RoboDK station: Vyankatesh_Robotic_Car_Painting_cell.rdk

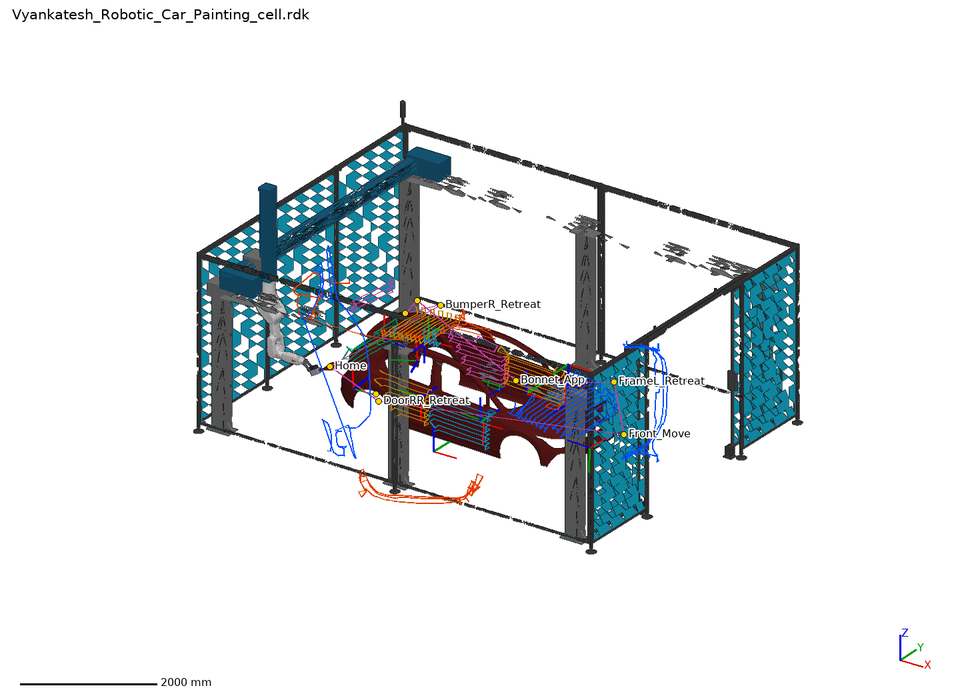
[picture v0: the station drawn from its stored meshes, robots at their saved joint values, targets as dots, program paths as lines]
Station Vyankatesh_Robotic_Car_Painting_cell (saved by RoboDK 6.1.1). Poses are relative to the parent item; angles as X-Y-Z fixed-axis rotations.
Station parameters (name, value as stored): Record_Record, 0, AttachCamera_Record, 0, Surface-Pattern-Generator-Settings, CollisionFreePlanner, ABB IRB 1300-10/1.15, CollisionFreePlanner-Rob ABB IRB 1300-10/1.15
  - frame Frame Car at (0, 0, 0) mm
    - object Trunk_T at (0, 0, 0) mm, size 559.9 x 1436.1 x 749.5 mm, geometry from Trunk_T.stl
    - object Bumper_F_T at (0, 0, 0) mm, size 772.5 x 1766.9 x 440.3 mm, geometry from Bumper_F_T.stl
    - object Bonnet_T at (0, 0, 0) mm, size 1078.9 x 1587.5 x 289.9 mm, geometry from Bonnet_T.stl
    - object Bumper_R_T at (0, 0, 0) mm, size 544.2 x 1726.4 x 536 mm, geometry from Bumper_R_T.stl
    - object Door_FL_T at (0, 0, 0) mm, size 1221.6 x 315.9 x 1113.7 mm, geometry from Door_FL_T.stl
    - object Door_FR_T at (0, 0, 0) mm, size 1221.6 x 316 x 1113.7 mm, geometry from Door_FR_T.stl
    - object Door_RL_T at (0, 0, 0) mm, size 1086.1 x 333.6 x 1090.9 mm, geometry from Door_RL_T.stl
    - object Door_RR_T at (0, 0, 0) mm, size 1086.1 x 333.6 x 1090.9 mm, geometry from Door_RR_T.stl
    - object Frame_T at (0, 0, 0) mm, size 3764.9 x 1786.8 x 1235.6 mm, geometry from Frame_T.stl
    - object Fuel_T at (0, 0, 0) mm, size 294.3 x 103.3 x 136.3 mm, geometry from Fuel_T.stl
    - object Top_T at (0, 0, 0) mm, size 810.7 x 1028.1 x 90.5 mm, geometry from Top_T.stl
    - frame Top2 at (-681.94, -447.22, 1360.45) mm, rotated rx -179.26 ry 1.08 rz -179.99 deg
    - frame Bonnet at (1052.19, 738.82, 942.03) mm, rotated rx 179.6 ry 0.01 rz 1.05 deg
    - frame DoorFL at (817.67, 994, 100.47) mm, rotated rx 105.9 ry -86.47 rz -19.07 deg
      - object DoorFL (SPG) at (0, 0, 0) mm
    - frame DoorRL at (-245.46, 977.17, 107.87) mm, rotated rx 13.73 ry -85.02 rz 76.6 deg
      - object DoorRL (SPG) at (0, 0, 0) mm
    - frame DoorFR at (798.13, -1053.51, 668.15) mm, rotated rx 42.25 ry 86.13 rz 132.32 deg
      - object DoorFR (SPG) at (0, 0, 0) mm
    - frame BumperF at (2280.3, -471.89, 411.2) mm, rotated rx -89.5 ry -0.21 rz 86.56 deg
    - frame DoorRR at (-287.77, -1076.71, 765.51) mm, rotated rx 87.83 ry 88.44 rz 179.37 deg
    - frame Bumper_R at (-1751.94, 908.52, 146.56) mm, rotated rx -73.11 ry -86.07 rz -175.08 deg
    - frame Trunk at (-2141.31, 613.21, 513.17) mm, rotated rx 88.99 ry -89.81 rz 85.05 deg
    - frame FrameL at (-1577.6, 957.23, 510.2) mm, rotated rx 93.66 ry 0 rz 0 deg
      - object FrameL (SPG) at (0, 0, 0) mm
    - frame FrameR at (-1577.79, -967.62, 493.6) mm, rotated rx 8.18 ry -85.7 rz -98.2 deg
      - object FrameR (SPG) at (0, 0, 0) mm
  - frame Cartesian Robot at (0, 0, 0) mm
    - robot My Mechanism: 3 axes
        modified DH rows (alpha deg, a mm, theta deg, d mm): 0, 0, 0, 0 linear; 90, 0, 90, 0 linear; 90, 0, 0, 0 linear
        base shift (0, 0, 0) mm, rotated rx 0 ry -90 rz 180 deg
        joint limits [0, -370, 0] to [5800, 3840, 1100]; home [0, 0, 0]; saved at [0, 0, 0]
      - robot ABB IRB 1300-10/1.15: 6 axes, payload 10 kg, reach 1150 mm, repeatability 0.023 mm, weight 78 kg
          modified DH rows (alpha deg, a mm, theta deg, d mm): 0, 0, 0, 544; -90, 150, -90, 0; 0, 575, 0, 0; -90, 40, 0, 425; 90, 0, 0, 0; -90, 0, 180, 90
          joint limits [-180, -95, -210, -230, -130, -400] to [180, 155, 65, 230, 130, 400]; home [0, 0, 0, 0, 0, 0]; saved at [0, 0, 0, 0, 0, 0]
        - tool Generic Paint Sprayer, TCP at (50, 0, 450) mm, rotated rx 0 ry 30 rz 0 deg, size 277.6 x 203.2 x 501.7 mm
  - frame Frame_Prog at (0, 0, 0) mm
    - target FrameL_Retreat (joint target) at (1421.65, 1379.32, 501.57) mm, rotated rx 178.9 ry 2.61 rz -172.87 deg; joints [31.932, 104.546, -125.413, -151.221, 47.063, 305.481, 2815.734, 3665.468, 738.344] of ABB IRB 1300-10/1.15
    - target Front_Move (Cartesian target) at (2873.26, -440.24, 778.86) mm, rotated rx 124.39 ry -0.68 rz -178.84 deg; joints [-120.26, 86.657, -7.45, -58.906, -114.481, 262.387, 5647.341, 170.911, 1082.66] of ABB IRB 1300-10/1.15
    - target Home (joint target) at (-1449.44, -1750.18, 1201) mm, rotated rx 0 ry -60 rz 180 deg; joints [0, 0, 0, 0, 0, 0, 0, 0, 0] of ABB IRB 1300-10/1.15
    - target BumperR_Retreat (joint target) at (-1695.61, 1414.09, 864.31) mm, rotated rx -107.53 ry 4.62 rz -165.7 deg; joints [-39.158, -91.932, 7.052, 83.863, 76.705, 97.807, 853.022, 3830.081, 364.531] of ABB IRB 1300-10/1.15
    - target Trunk_App (Cartesian target) at (-2045.19, 1025.35, 789.85) mm, rotated rx 93.3 ry 0.38 rz 73.69 deg; joints [-81.249, 102.661, -200.517, 127.066, 82.558, -85.71, 17.635, 2525.27, 659.745] of ABB IRB 1300-10/1.15
    - target Top_Retreat (joint target) at (-1442.79, 464.8, 1389.13) mm, rotated rx -170.97 ry 7.12 rz -173.76 deg; joints [13.22, 135.95, -182.37, -143.59, 7.01, 303.87, 37.44, 2446.95, 0] of ABB IRB 1300-10/1.15
    - target Bonnet_App (joint target) at (1119.24, -686.1, 1265.98) mm, rotated rx 177.3 ry -5.95 rz 179.99 deg; joints [172.493, 123.347, -162.887, -179.232, 74.635, 188.011, 4433.831, 1162.767, 1.741] of ABB IRB 1300-10/1.15
    - target DoorRR_Retreat (joint target) at (-794.82, -1444.65, 696.6) mm, rotated rx 75.81 ry -0.27 rz 178.92 deg; joints [-164.383, 16.979, -25.325, 79.856, 107.569, -167.519, 2238.906, -364.928, 537.904] of ABB IRB 1300-10/1.15
    - target FrameR_App (Cartesian target) at (-1034.25, -1174.19, 640.35) mm, rotated rx 101.61 ry -1.74 rz -171.59 deg; joints [-36.204, 78.94, -160.975, 146.937, -72.367, 90.08, 787.656, -367.42, 482.946] of ABB IRB 1300-10/1.15
  - machining project FrameR: rotZ(0) | rotz(0) | onStart | onPathStart | onApproach | onPoint | onRetract | onFinish | SetRPM(%1) | SetTool(%1) | Extruder(%1) | default | default | OutOnMov(%1) | OutOffMov(%1) | onPathFinish | M_RunCode(%1)
  - machining project FrameL: rotZ(0) | rotz(0) | onStart | onPathStart | onApproach | onPoint | onRetract | onFinish | SetRPM(%1) | SetTool(%1) | Extruder(%1) | default | default | OutOnMov(%1) | OutOffMov(%1) | onPathFinish | M_RunCode(%1)
  - machining project BumperF: rotZ(0) | rotz(0) | onStart | onPathStart | onApproach | onPoint | onRetract | onFinish | SetRPM(%1) | SetTool(%1) | Extruder(%1) | default | default | OutOnMov(%1) | OutOffMov(%1) | onPathFinish | M_RunCode(%1)
  - machining project Bonnet: rotZ(0) | onStart | onPathStart | onApproach | onPoint | onRetract | onFinish | SetRPM(%1) | SetTool(%1) | Extruder(%1) | default | default | OutOnMov(%1) | OutOffMov(%1) | onPathFinish | M_RunCode(%1)
  - machining project Top2: rotZ(0) | rotZ(0) | onStart | onPathStart | onApproach | onPoint | onRetract | onFinish | SetRPM(%1) | SetTool(%1) | Extruder(%1) | default | default | OutOnMov(%1) | OutOffMov(%1) | onPathFinish | M_RunCode(%1)
  - machining project DoorFL: rotZ(0) | rotz(0) | onStart | onPathStart | onApproach | onPoint | onRetract | onFinish | SetRPM(%1) | SetTool(%1) | Extruder(%1) | default | default | OutOnMov(%1) | OutOffMov(%1) | onPathFinish | M_RunCode(%1)
  - machining project DoorRL: rotZ(0) | rotz(0) | onStart | onPathStart | onApproach | onPoint | onRetract | onFinish | SetRPM(%1) | SetTool(%1) | Extruder(%1) | default | default | OutOnMov(%1) | OutOffMov(%1) | onPathFinish | M_RunCode(%1)
  - machining project DoorFR: rotZ(0) | rotZ(0) | onStart | onPathStart | onApproach | onPoint | onRetract | onFinish | SetRPM(%1) | SetTool(%1) | Extruder(%1) | default | default | OutOnMov(%1) | OutOffMov(%1) | onPathFinish | M_RunCode(%1)
  - machining project DoorRR: rotZ(0) | rotz(0) | onStart | onPathStart | onApproach | onPoint | onRetract | onFinish | SetRPM(%1) | SetTool(%1) | Extruder(%1) | default | default | OutOnMov(%1) | OutOffMov(%1) | onPathFinish | M_RunCode(%1)
  - machining project Trunk: rotZ(0) | rotz(0) | onStart | onPathStart | onApproach | onPoint | onRetract | onFinish | SetRPM(%1) | SetTool(%1) | Extruder(%1) | default | default | OutOnMov(%1) | OutOffMov(%1) | onPathFinish | M_RunCode(%1)
  - machining project Bumper_R: rotZ(0) | rotz(0) | onStart | onPathStart | onApproach | onPoint | onRetract | onFinish | SetRPM(%1) | SetTool(%1) | Extruder(%1) | default | default | OutOnMov(%1) | OutOffMov(%1) | onPathFinish | M_RunCode(%1)
  - program Bonnet (314 instructions, listed below)
  - program Top2 (192 instructions, listed below)
  - program DoorRR_C (126 instructions, listed below)
  - program DoorRL_C (142 instructions, listed below)
  - program DoorFL_C (149 instructions, listed below)
  - program DoorFR_C (147 instructions, listed below)
  - program DoorFR (14 instructions, listed below)
  - program BumperR_C (354 instructions, listed below)
  - program Trunk_C (101 instructions, listed below)
  - program Trunk_Top_C (58 instructions, listed below)
  - program Top2_C (192 instructions, listed below)
  - program BumperF (415 instructions, listed below)
  - program BumperF_C (415 instructions, listed below)
  - program FrameL_C (243 instructions, listed below)
  - program FrameR_C (273 instructions, listed below)
  - program Main_Prog (22 instructions, listed below)
  - frame Cell  at (0, 0, 0) mm
    - frame Left at (0, -1180, 0) mm
      - object LeftGlass at (0, 0, 0) mm, size 6 x 1164 x 2469 mm, geometry from LeftGlass.stl
      - object LeftGlassFrame at (0, 0, 0) mm, size 172 x 1253 x 2620 mm, geometry from LeftGlassFrame.stl
    - frame Right at (0, 1180, 0) mm
      - object RightGlass at (0, 0, 0) mm, size 6 x 1166 x 2471 mm, geometry from RightGlass.stl
      - object RightGlassFrame at (0, 0, 0) mm, size 172 x 1253 x 2620 mm, geometry from RightGlassFrame.stl
  - object Floor at (0, 0, 0) mm, size 8000 x 5600 x 0 mm, geometry from Floor.stl
  - object OuterGlass at (0, 0, 0) mm, size 7005.9 x 5255.9 x 2661 mm, geometry from OuterGlass.stl
  - object GlassFrame at (0, 0, 0) mm, size 7159.9 x 5409.9 x 3270 mm, geometry from GlassFrame.stl
  - program DoorRR (126 instructions, listed below)
  - program FrameL (45 instructions, listed below)
  - program FrameR (273 instructions, listed below)
  - program DoorFL (22 instructions, listed below)
  - program DoorRL (15 instructions, listed below)
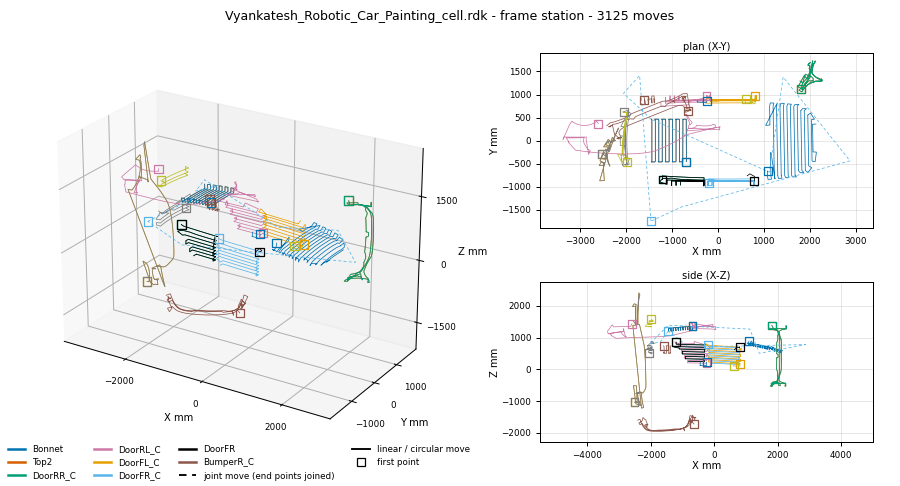
[picture p0: tool path of Vyankatesh_Robotic_Car_Painting_cell.rdk in frame station, 3125 of 3125 moves have a stored position in this frame; points joined in program order, loops and branches not executed]

--- program Bonnet (robot ABB IRB 1300-10/1.15) ---
  Smooth(1)
  Set speed (1000.0 mm/s)
  Set Ref.: Bonnet
  Set Tool: Generic Paint Sprayer
  Show Generic Paint Sprayer
  MoveJ 1 to (13.71, 1405.55, 66.05) mm, rotated rx -3.07 ry 7.94 rz -179.16 deg; joints [173.742, 90.77, -145.127, -180, 57.846, 186.984, 4434.016, 1162.706, 0.414]
  MoveL 2 to (13.71, 1405.55, 66.05) mm, rotated rx -3.07 ry 7.94 rz -179.16 deg; joints [173.742, 90.77, -145.127, -180, 57.846, 186.984, 4434.017, 1162.706, 0.414]
  MoveL 3 to (0, 1400, 164.95) mm, rotated rx -3.07 ry 7.94 rz -179.16 deg; joints [173.742, 90.769, -145.127, -180, 57.846, 186.984, 4420.212, 1167.307, 99.349]
  MoveL 4 to (0, 1400, 164.95) mm, rotated rx -3.07 ry 7.94 rz -179.16 deg; joints [173.742, 90.769, -145.127, -180, 57.846, 186.984, 4420.212, 1167.307, 99.349]
  Set speed (200.0 mm/s)
  MoveL 5 to (0, 1500, 204.66) mm, rotated rx -53.96 ry 9.04 rz 178.26 deg; joints [162.372, 90.769, -145.127, -214.939, 81.944, 234.484, 4381.306, 868.259, 332.309]
  Set speed (1000.0 mm/s)
  MoveL 6 to (0, 1500, 204.66) mm, rotated rx -53.96 ry 9.04 rz 178.26 deg; joints [162.372, 90.769, -145.127, -214.939, 81.944, 234.484, 4381.306, 868.259, 332.309]
  MoveL 7 to (11.7, 1580.54, 146.56) mm, rotated rx -53.96 ry 9.04 rz 178.26 deg; joints [162.372, 90.77, -145.127, -214.939, 81.944, 234.484, 4394.48, 788.358, 273.639]
  Set speed (1000.0 mm/s)
  MoveL 8 to (86.8, 1577.85, 157.52) mm, rotated rx -51.38 ry 9.02 rz 178.52 deg; joints [163.545, 90.769, -145.127, -214.254, 79.866, 232.519, 4475.298, 788.36, 267.392]
  MoveL 9 to (75, 1500, 219.17) mm, rotated rx -51.38 ry 9.02 rz 178.52 deg; joints [163.545, 90.769, -145.127, -214.254, 79.866, 232.519, 4462.081, 865.544, 329.584]
  MoveL 10 to (75, 1500, 219.17) mm, rotated rx -51.38 ry 9.02 rz 178.52 deg; joints [163.545, 90.769, -145.127, -214.254, 79.866, 232.519, 4462.081, 865.544, 329.584]
  Set speed (200.0 mm/s)
  MoveL 11 to (75, 1400, 175.28) mm, rotated rx -2.63 ry 8.05 rz -179.16 deg; joints [163.545, 106.008, -145.127, -175.627, 72.598, 194.93, 4527.686, 1355.214, 329.584]
  MoveL 12 to (75, 1300, 170.07) mm, rotated rx -3.56 ry 8.28 rz -179.19 deg; joints [164.42, 106.008, -145.153, -176.848, 72.598, 194.93, 4532.073, 1432.375, 324.681]
  MoveL 13 to (75, 1200, 162.92) mm, rotated rx -2 ry 7.25 rz -179.12 deg; joints [166.99, 106.008, -145.153, -176.244, 73.416, 191.618, 4532.073, 1502.111, 320.532]
  MoveL 14 to (75, 1100, 159.11) mm, rotated rx -1.73 ry 6.88 rz -179.11 deg; joints [167.767, 106.008, -145.153, -176.244, 73.775, 190.768, 4529.877, 1591.137, 318.443]
  MoveL 15 to (75, 1000, 155.9) mm, rotated rx -1.44 ry 7.2 rz -179.12 deg; joints [167.77, 106.24, -145.152, -176.048, 73.647, 190.576, 4531.483, 1693.74, 318.443]
  Set speed (1000.0 mm/s)
  MoveL 16 to (75, 1000, 155.9) mm, rotated rx -1.44 ry 7.2 rz -179.12 deg; joints [167.77, 106.24, -145.152, -176.048, 73.647, 190.576, 4531.483, 1693.74, 318.443]
  MoveL 17 to (87.48, 1002.7, 56.72) mm, rotated rx -1.44 ry 7.2 rz -179.12 deg; joints [167.77, 106.24, -145.152, -176.048, 73.647, 190.576, 4544.012, 1691.978, 219.247]
  Set speed (1000.0 mm/s)
  MoveL 18 to (163.33, 1574.44, 167.94) mm, rotated rx -44.22 ry 24.07 rz -167.42 deg; joints [161.786, 90.814, -145.127, -206.546, 69.381, 247.678, 4571.543, 889.471, 203.361]
  MoveL 19 to (150, 1500, 233.37) mm, rotated rx -44.22 ry 24.07 rz -167.42 deg; joints [161.786, 90.814, -145.127, -206.546, 69.382, 247.678, 4556.853, 963.186, 269.318]
  MoveL 20 to (150, 1500, 233.37) mm, rotated rx -44.22 ry 24.07 rz -167.42 deg; joints [161.786, 90.814, -145.127, -206.546, 69.382, 247.678, 4556.853, 963.186, 269.318]
  Set speed (200.0 mm/s)
  MoveL 21 to (150, 1400, 185.67) mm, rotated rx 0.71 ry 8.41 rz -158.95 deg; joints [180, 101.307, -145.127, -171.069, 66.652, 194.666, 4644.083, 1152.192, 269.318]
  MoveL 22 to (150, 1300, 180.88) mm, rotated rx -8.15 ry 4.46 rz 140.73 deg; joints [127.726, 83.623, -166.891, -182.813, 33.065, 197.095, 4139.747, 1597.912, 0.019]
  MoveL 23 to (150, 1200, 172.83) mm, rotated rx -2.4 ry 7.56 rz -179.14 deg; joints [25.975, 87.43, -169.901, -43.466, 16.467, 198.768, 2962.972, 1597.586, 18.083]
  MoveL 24 to (150, 1100, 168.79) mm, rotated rx -2.16 ry 7.38 rz -179.13 deg; joints [25.908, 87.621, -170.162, -42.349, 16.618, 197.63, 2959.562, 1698.654, 17.072]
  MoveL 25 to (150, 1000, 165.32) mm, rotated rx -1.64 ry 7.21 rz -179.12 deg; joints [25.707, 87.861, -170.491, -40.208, 16.705, 195.488, 2955.557, 1800.56, 17.072]
  MoveL 26 to (150, 900, 162.41) mm, rotated rx -1.26 ry 7.12 rz -179.12 deg; joints [25.558, 88.036, -170.732, -38.697, 16.743, 193.978, 2952.499, 1901.9, 16.797]
  MoveL 27 to (150, 800, 160.25) mm, rotated rx -1.02 ry 6.68 rz -179.11 deg; joints [25.455, 88.057, -170.76, -37.493, 17.124, 192.798, 2946.147, 2002.771, 16.797]
  MoveL 28 to (150, 700, 159.04) mm, rotated rx 0.41 ry 7.43 rz -179.12 deg; joints [24.734, 88.057, -170.76, -32.755, 16.105, 188.203, 2947.144, 2106.644, 14.156]
  MoveL 29 to (150, 600, 159.34) mm, rotated rx 0.28 ry 6.68 rz -179.12 deg; joints [24.734, 87.748, -170.76, -32.228, 17.13, 187.718, 2940.681, 2204.426, 14.157]
  MoveL 30 to (150, 500, 160.27) mm, rotated rx 0.78 ry 7.01 rz -179.12 deg; joints [24.474, 87.675, -170.719, -30.467, 16.76, 186.011, 2940.681, 2305.628, 14.157]
  MoveL 31 to (150, 400, 161.65) mm, rotated rx 0.99 ry 7.45 rz -179.12 deg; joints [24.363, 87.589, -170.601, -29.905, 16.266, 185.477, 2942.074, 2406.202, 14.157]
  MoveL 32 to (150, 300, 163.74) mm, rotated rx 1.37 ry 7.2 rz -179.12 deg; joints [24.17, 87.589, -170.601, -28.388, 16.481, 184.008, 2936.908, 2507.18, 17.764]
  MoveL 33 to (150, 200, 169.2) mm, rotated rx 2.84 ry 8.35 rz -179.06 deg; joints [23.441, 87.248, -170.135, -23.017, 15.142, 178.814, 2940.939, 2611.654, 17.919]
  MoveL 34 to (150, 100, 172.42) mm, rotated rx 1.6 ry 7.77 rz -179.1 deg; joints [23.441, 86.759, -170.135, -26.264, 16.178, 182.487, 2937.523, 2699.259, 17.919]
  MoveL 35 to (150, 0, 193.42) mm, rotated rx 48.1 ry 9.85 rz -176.1 deg; joints [6.576, 86.759, -170.136, 60.139, 45.852, 96.029, 2889.461, 2951.486, 197.833]
  Set speed (1000.0 mm/s)
  MoveL 36 to (150, 0, 193.42) mm, rotated rx 48.1 ry 9.85 rz -176.1 deg; joints [6.576, 86.759, -170.136, 60.139, 45.852, 96.029, 2889.461, 2951.486, 197.833]
  MoveL 37 to (166.47, -73.48, 127.62) mm, rotated rx 48.1 ry 9.85 rz -176.1 deg; joints [6.576, 86.759, -170.136, 60.139, 45.852, 96.029, 2904.579, 3025.719, 132.557]
  Set speed (1000.0 mm/s)
  MoveL 38 to (89.54, -78.19, 114.09) mm, rotated rx 52.11 ry 9.16 rz -176.52 deg; joints [5.072, 86.759, -170.136, 61.133, 49.725, 94.485, 2815.202, 3031.106, 147.378]
  MoveL 39 to (75, 0, 174.71) mm, rotated rx 52.11 ry 9.16 rz -176.52 deg; joints [5.072, 86.759, -170.136, 61.133, 49.725, 94.486, 2802.092, 2952.242, 207.449]
  MoveL 40 to (75, 0, 174.71) mm, rotated rx 52.11 ry 9.16 rz -176.52 deg; joints [5.072, 86.759, -170.136, 61.133, 49.725, 94.486, 2802.092, 2952.242, 207.449]
  Set speed (200.0 mm/s)
  MoveL 41 to (75, 100, 161.89) mm, rotated rx 1.85 ry 8.11 rz -179.09 deg; joints [23.489, 88.002, -170.136, -27.629, 14.727, 183.787, 2856.802, 2704.635, 19.313]
  MoveL 42 to (75, 200, 158.17) mm, rotated rx 2.73 ry 8.3 rz -179.07 deg; joints [23.489, 88.444, -170.136, -25.354, 14.108, 181.209, 2857.15, 2613.667, 19.312]
  MoveL 43 to (75, 300, 153.75) mm, rotated rx 1.3 ry 7.73 rz -179.11 deg; joints [24.186, 88.444, -170.136, -31.197, 14.806, 186.915, 2857.632, 2509.61, 15.205]
  MoveL 44 to (75, 400, 153.25) mm, rotated rx -65.18 ry 32.47 rz -81.47 deg; joints [-7.384, 82.47, -173.542, 30.828, 55.97, 290.824, 2599.504, 2142.82, 179.665]
  Set speed (1000.0 mm/s)
  MoveL 45 to (75, 400, 153.25) mm, rotated rx -65.18 ry 32.47 rz -81.47 deg; joints [-7.384, 82.47, -173.542, 30.828, 55.97, 290.824, 2599.504, 2142.82, 179.665]
  MoveL 46 to (-18.1, 408.83, 117.84) mm, rotated rx -48.18 ry -57.92 rz -132.58 deg; joints [5.789, 76.051, -169.247, 0, 99.953, 203.081, 2424.003, 2179.227, 396.057]
  Set speed (1000.0 mm/s)
  MoveL 47 to (242.54, -75.07, 148.77) mm, rotated rx 49.67 ry 10.26 rz -175.45 deg; joints [5.789, 76.051, -169.247, 55.04, 52.306, 105.502, 3073.622, 3019.948, 61.16]
  MoveL 48 to (225, 0, 212.46) mm, rotated rx 49.67 ry 10.26 rz -175.45 deg; joints [5.789, 76.051, -169.247, 55.04, 52.306, 105.502, 3057.455, 2944.119, 124.315]
  MoveL 49 to (225, 0, 212.46) mm, rotated rx 49.67 ry 10.26 rz -175.45 deg; joints [5.789, 76.051, -169.247, 55.04, 52.306, 105.502, 3057.455, 2944.119, 124.315]
  Set speed (200.0 mm/s)
  MoveL 50 to (225, 100, 183.39) mm, rotated rx 0.83 ry 8.18 rz -179.11 deg; joints [15.296, 83.487, -177.068, -10.85, 25.36, 174.895, 3057.454, 2574.979, 0]
  MoveL 51 to (225, 200, 180.77) mm, rotated rx 2.66 ry 8.52 rz -179.06 deg; joints [15.296, 83.901, -177.068, -7.153, 24.807, 170.698, 3058.945, 2491.778, 0]
  MoveL 52 to (225, 300, 173.64) mm, rotated rx 1.36 ry 7.35 rz -179.12 deg; joints [15.88, 84.388, -177.768, -10.555, 26.023, 173.843, 3053.064, 2386.704, 0]
  MoveL 53 to (225, 400, 171.5) mm, rotated rx 1.18 ry 7.79 rz -179.11 deg; joints [16.011, 84.85, -177.768, -11.109, 25.117, 174.348, 3055.565, 2287.744, 0]
  MoveL 54 to (225, 500, 169.85) mm, rotated rx 0.84 ry 7.43 rz -179.12 deg; joints [16.182, 84.988, -177.967, -12.016, 25.501, 175.176, 3055.056, 2186.543, 0]
  MoveL 55 to (225, 600, 168.94) mm, rotated rx 0.53 ry 7.14 rz -179.12 deg; joints [16.33, 85.067, -178.08, -12.799, 25.81, 175.895, 3054.866, 2085.487, 0]
  MoveL 56 to (225, 700, 168.3) mm, rotated rx 0.46 ry 7.35 rz -179.12 deg; joints [16.389, 85.287, -178.08, -13.055, 25.373, 176.127, 3057.115, 1986.104, 0]
  MoveL 57 to (225, 800, 169.49) mm, rotated rx -1.24 ry 7.12 rz -179.12 deg; joints [17.175, 85.179, -177.924, -17.239, 25.498, 180.034, 3059.26, 1880.248, 0]
  MoveL 58 to (225, 900, 171.99) mm, rotated rx -1.33 ry 6.99 rz -179.12 deg; joints [17.227, 85.28, -177.924, -17.522, 25.536, 180.297, 3059.26, 1780.347, 3.097]
  MoveL 59 to (225, 1000, 174.93) mm, rotated rx -1.68 ry 7.42 rz -179.13 deg; joints [17.384, 85.177, -177.776, -18.423, 25.066, 181.15, 3065.255, 1679.079, 3.097]
  MoveL 60 to (225, 1100, 178.7) mm, rotated rx -2.17 ry 8.02 rz -179.15 deg; joints [17.597, 85.034, -177.569, -19.725, 24.409, 182.385, 3072.997, 1577.25, 3.097]
  MoveL 61 to (225, 1200, 182.76) mm, rotated rx -2.2 ry 7.73 rz -179.14 deg; joints [17.603, 85.034, -177.569, -19.748, 24.7, 182.411, 3072.215, 1477.151, 7.244]
  MoveL 62 to (225, 1300, 192.42) mm, rotated rx -2.69 ry 8.46 rz -179.18 deg; joints [17.714, 84.444, -176.724, -21.177, 23.751, 183.883, 3079.788, 1374.447, 8.221]
  MoveL 63 to (225, 1400, 196.36) mm, rotated rx -1.65 ry 8.59 rz -179.16 deg; joints [17.714, 84.583, -176.724, -19.035, 23.457, 181.445, 3081.636, 1283.763, 12.105]
  MoveL 64 to (225, 1500, 247.21) mm, rotated rx -41.7 ry 9.43 rz 178.83 deg; joints [27.955, 71.742, -159.319, -88.579, 43.502, 254.167, 3123.032, 976.712, 51.789]
  Set speed (1000.0 mm/s)
  MoveL 65 to (225, 1500, 247.21) mm, rotated rx -41.7 ry 9.43 rz 178.83 deg; joints [27.955, 71.742, -159.319, -88.579, 43.502, 254.167, 3123.032, 976.712, 51.789]
  MoveL 66 to (238.58, 1566.25, 173.55) mm, rotated rx -41.7 ry 9.43 rz 178.83 deg; joints [29.173, 74.127, -159.319, -92.303, 43.597, 257.628, 3123.032, 935.899, 0]
  Set speed (1000.0 mm/s)
  MoveL 67 to (315.52, 1560.78, 183.61) mm, rotated rx -37.7 ry 10.16 rz 178.53 deg; joints [27.986, 75.504, -159.319, -92.621, 39.841, 257.853, 3190.269, 962.686, 0]
  MoveL 68 to (300, 1500, 261.49) mm, rotated rx -37.7 ry 10.16 rz 178.53 deg; joints [27.986, 75.504, -159.319, -92.621, 39.841, 257.853, 3173.641, 1022.617, 78.302]
  MoveL 69 to (300, 1500, 261.49) mm, rotated rx -37.7 ry 10.16 rz 178.53 deg; joints [27.986, 75.504, -159.319, -92.621, 39.841, 257.853, 3173.641, 1022.617, 78.302]
  Set speed (200.0 mm/s)
  MoveL 70 to (300, 1400, 208.07) mm, rotated rx -1.39 ry 8.99 rz -179.17 deg; joints [17.09, 87.326, -175.277, -21.576, 19.105, 184.796, 3126.615, 1290.083, 47.242]
  MoveL 71 to (300, 1300, 204.58) mm, rotated rx -2.31 ry 9.55 rz -179.22 deg; joints [16.15, 87.326, -175.277, -23.211, 18.622, 187.649, 3126.615, 1371.082, 43.238]
  MoveL 72 to (300, 1200, 193.84) mm, rotated rx -2.35 ry 8.91 rz -179.19 deg; joints [16.15, 87.762, -175.895, -22.88, 19.432, 187.336, 3120.036, 1470.451, 39.287]
  MoveL 73 to (300, 1100, 189.49) mm, rotated rx -2.12 ry 8.59 rz -179.17 deg; joints [16.081, 88.023, -176.265, -21.971, 19.824, 186.418, 3115.771, 1571.51, 39.081]
  MoveL 74 to (300, 1000, 185.81) mm, rotated rx -1.83 ry 8.63 rz -179.17 deg; joints [15.939, 88.053, -176.308, -21.088, 19.772, 185.583, 3113.884, 1672.287, 36.248]
  MoveL 75 to (300, 900, 182.49) mm, rotated rx -1.49 ry 8.68 rz -179.16 deg; joints [15.765, 88.088, -176.358, -19.999, 19.711, 184.554, 3111.995, 1773.235, 33.807]
  MoveL 76 to (300, 800, 179.69) mm, rotated rx -1.28 ry 8.26 rz -179.15 deg; joints [15.674, 88.189, -176.502, -19.237, 20.15, 183.816, 3106.38, 1873.929, 33.807]
  MoveL 77 to (300, 700, 178.51) mm, rotated rx 0.42 ry 8.27 rz -179.11 deg; joints [14.803, 88.236, -176.569, -13.977, 20.124, 178.867, 3101.896, 1978.338, 33.807]
  MoveL 78 to (300, 600, 179.27) mm, rotated rx 0.66 ry 8.76 rz -179.1 deg; joints [14.68, 88.216, -176.54, -13.21, 19.632, 178.149, 3104.063, 2078.956, 33.807]
  MoveL 79 to (300, 500, 180.56) mm, rotated rx 1.01 ry 8.7 rz -179.09 deg; joints [14.502, 88.216, -176.54, -12.117, 19.701, 177.121, 3101.147, 2179.85, 36.013]
  MoveL 80 to (300, 400, 182.21) mm, rotated rx 1.26 ry 8.59 rz -179.09 deg; joints [14.374, 88.216, -176.54, -11.346, 19.823, 176.394, 3097.913, 2280.477, 38.718]
  MoveL 81 to (300, 300, 184.43) mm, rotated rx 1.56 ry 9.04 rz -179.07 deg; joints [14.207, 88.036, -176.285, -10.336, 19.316, 175.463, 3099.179, 2381.233, 38.718]
  MoveL 82 to (300, 200, 192.84) mm, rotated rx 2.59 ry 9.4 rz -179.02 deg; joints [13.689, 87.953, -176.21, -6.909, 19.057, 172.229, 3099.179, 2484.02, 46.473]
  MoveL 83 to (300, 100, 194.82) mm, rotated rx 0.83 ry 9.24 rz -179.09 deg; joints [13.689, 87.711, -176.211, -11.528, 19.32, 177.395, 3097.796, 2568.243, 46.707]
  MoveL 84 to (300, 0, 232.6) mm, rotated rx 41.6 ry 10.8 rz -175.86 deg; joints [-6.021, 87.711, -176.211, 68.056, 42.901, 105.13, 3088.96, 2757.637, 205.756]
  Set speed (1000.0 mm/s)
  MoveL 85 to (300, 0, 232.6) mm, rotated rx 41.6 ry 10.8 rz -175.86 deg; joints [-6.021, 87.711, -176.211, 68.056, 42.901, 105.13, 3088.96, 2757.637, 205.756]
  MoveL 86 to (318.77, -65.21, 159.15) mm, rotated rx 41.6 ry 10.8 rz -175.86 deg; joints [-6.021, 87.711, -176.211, 68.056, 42.901, 105.13, 3106.537, 2823.697, 132.769]
  Set speed (1000.0 mm/s)
  MoveL 87 to (394.09, -63.48, 176.58) mm, rotated rx 40.3 ry 10.95 rz -175.88 deg; joints [-5.321, 87.766, -176.211, 67.069, 41.703, 105.865, 3182.413, 2823.062, 143.079]
  MoveL 88 to (375, 0, 251.46) mm, rotated rx 40.3 ry 10.95 rz -175.88 deg; joints [-5.321, 87.766, -176.211, 67.069, 41.703, 105.865, 3164.491, 2758.721, 217.504]
  MoveL 89 to (375, 0, 251.46) mm, rotated rx 40.3 ry 10.95 rz -175.88 deg; joints [-5.321, 87.766, -176.211, 67.069, 41.703, 105.865, 3164.491, 2758.721, 217.504]
  Set speed (200.0 mm/s)
  MoveL 90 to (375, 100, 207.39) mm, rotated rx 0.55 ry 10.1 rz -179.09 deg; joints [13.83, 87.766, -176.211, -12.371, 18.395, 178.193, 3180.679, 2568.934, 57.639]
  MoveL 91 to (375, 200, 205.89) mm, rotated rx 2.6 ry 10.23 rz -178.98 deg; joints [13.83, 88.078, -176.211, -6.727, 18.114, 171.926, 3181.211, 2487.437, 58.72]
  MoveL 92 to (375, 300, 196.95) mm, rotated rx 1.57 ry 9.8 rz -179.05 deg; joints [14.354, 88.197, -176.38, -10.315, 18.496, 175.304, 3181.025, 2384.58, 50.941]
  MoveL 93 to (375, 400, 194.55) mm, rotated rx 1.23 ry 9.65 rz -179.07 deg; joints [14.527, 88.254, -176.38, -11.497, 18.564, 176.419, 3181.65, 2283.834, 48.647]
  MoveL 94 to (375, 500, 192.59) mm, rotated rx 1 ry 9.63 rz -179.08 deg; joints [14.644, 88.254, -176.38, -12.262, 18.582, 177.14, 3183.59, 2183.241, 45.99]
  MoveL 95 to (375, 600, 191.19) mm, rotated rx 0.68 ry 9.25 rz -179.1 deg; joints [14.825, 88.373, -176.549, -13.366, 19, 178.164, 3182.849, 2082.442, 45.99]
  MoveL 96 to (375, 700, 190.31) mm, rotated rx 0.61 ry 9.24 rz -179.1 deg; joints [14.859, 88.373, -176.549, -13.585, 19.005, 178.369, 3184.727, 1982.29, 44.406]
  MoveL 97 to (375, 800, 191.51) mm, rotated rx -1.47 ry 9.25 rz -179.17 deg; joints [15.931, 88.325, -176.482, -20.389, 19.038, 184.772, 3190.004, 1876.825, 44.405]
  MoveL 98 to (375, 900, 194.48) mm, rotated rx -1.72 ry 9.6 rz -179.19 deg; joints [16.032, 88.185, -176.282, -21.327, 18.652, 185.686, 3195.013, 1775.96, 44.405]
  MoveL 99 to (375, 1000, 197.95) mm, rotated rx -1.86 ry 9.61 rz -179.2 deg; joints [16.097, 88.151, -176.234, -21.797, 18.641, 186.135, 3197.071, 1675.545, 46.812]
  MoveL 100 to (375, 1100, 202) mm, rotated rx -2.39 ry 10.09 rz -179.24 deg; joints [16.322, 87.923, -175.91, -23.8, 18.139, 188.075, 3203.415, 1573.734, 46.812]
  MoveL 101 to (375, 1200, 206.54) mm, rotated rx -2.44 ry 9.79 rz -179.23 deg; joints [16.352, 87.923, -175.91, -23.845, 18.441, 188.115, 3202.619, 1473.638, 51.377]
  MoveL 102 to (375, 1300, 217.6) mm, rotated rx -2.03 ry 10.57 rz -179.24 deg; joints [16.352, 87.453, -175.243, -23.259, 17.441, 187.396, 3210.369, 1377.45, 54.97]
  MoveL 103 to (375, 1400, 221) mm, rotated rx -1.2 ry 10.41 rz -179.19 deg; joints [16.352, 87.508, -175.243, -20.821, 17.466, 184.706, 3210.369, 1284.858, 58.398]
  MoveL 104 to (375, 1500, 276.56) mm, rotated rx -29.1 ry 11.25 rz 178.58 deg; joints [25.924, 79.147, -163.83, -87.251, 31.923, 250.899, 3248.664, 1064.43, 86.696]
  Set speed (1000.0 mm/s)
  MoveL 105 to (375, 1500, 276.56) mm, rotated rx -29.1 ry 11.25 rz 178.58 deg; joints [25.924, 79.147, -163.83, -87.251, 31.923, 250.899, 3248.664, 1064.43, 86.696]
  MoveL 106 to (393.24, 1548.2, 190.86) mm, rotated rx -29.1 ry 11.25 rz 178.58 deg; joints [25.924, 79.147, -163.83, -87.251, 31.923, 250.899, 3267.782, 1017.182, 0.665]
  Set speed (1000.0 mm/s)
  MoveL 107 to (470.75, 1541.56, 204.5) mm, rotated rx -24.91 ry 12.47 rz 178.4 deg; joints [24.056, 79.641, -163.83, -85.84, 27.687, 249.752, 3343.92, 1038.3, 0.665]
  MoveL 108 to (450, 1500, 293.05) mm, rotated rx -24.91 ry 12.47 rz 178.4 deg; joints [24.056, 79.64, -163.83, -85.838, 27.687, 249.75, 3322.418, 1078.84, 89.502]
  MoveL 109 to (450, 1500, 293.05) mm, rotated rx -24.91 ry 12.47 rz 178.4 deg; joints [24.056, 79.64, -163.83, -85.838, 27.687, 249.75, 3322.418, 1078.84, 89.502]
  Set speed (200.0 mm/s)
  MoveL 110 to (450, 1400, 235.27) mm, rotated rx -1.57 ry 11.98 rz -179.25 deg; joints [16.298, 86.244, -172.78, -24.148, 14.832, 188.239, 3291.716, 1284.532, 56.208]
  MoveL 111 to (450, 1300, 231.88) mm, rotated rx -2.49 ry 10.96 rz -179.29 deg; joints [16.298, 86.268, -172.814, -26.537, 15.986, 190.936, 3280.502, 1376.523, 56.208]
  MoveL 112 to (450, 1200, 220.89) mm, rotated rx -2.79 ry 11.21 rz -179.32 deg; joints [16.171, 86.268, -172.814, -27.528, 15.785, 192.139, 3280.58, 1472.42, 45.456]
  MoveL 113 to (450, 1100, 215.84) mm, rotated rx -2.44 ry 10.78 rz -179.28 deg; joints [16.073, 86.612, -173.293, -25.8, 16.274, 190.404, 3275.148, 1574.119, 45.456]
  MoveL 114 to (450, 1000, 211.48) mm, rotated rx -2.12 ry 10.68 rz -179.25 deg; joints [15.943, 86.743, -173.476, -24.509, 16.367, 189.139, 3272.269, 1675.333, 43.277]
  MoveL 115 to (450, 900, 207.67) mm, rotated rx -1.59 ry 10.35 rz -179.21 deg; joints [15.732, 86.986, -173.816, -22.34, 16.711, 187.012, 3267.276, 1777.314, 43.277]
  MoveL 116 to (450, 800, 204.58) mm, rotated rx -1.69 ry 10.65 rz -179.22 deg; joints [15.718, 86.986, -173.816, -22.76, 16.419, 187.472, 3268.202, 1876.273, 40.202]
  MoveL 117 to (450, 700, 203.34) mm, rotated rx 0.81 ry 10.66 rz -179.07 deg; joints [14.541, 87.041, -173.892, -13.488, 16.297, 178.578, 3262.711, 1984.048, 40.202]
  MoveL 118 to (450, 600, 204.37) mm, rotated rx 0.72 ry 10.35 rz -179.08 deg; joints [14.542, 86.792, -173.892, -13.596, 16.843, 178.705, 3260.003, 2082.718, 40.219]
  MoveL 119 to (450, 500, 205.98) mm, rotated rx 1.23 ry 10.65 rz -179.04 deg; joints [14.298, 86.674, -173.753, -11.727, 16.545, 176.92, 3260.003, 2184.256, 40.766]
  MoveL 120 to (450, 400, 208.16) mm, rotated rx 1.57 ry 10.79 rz -179.02 deg; joints [14.14, 86.622, -173.753, -10.42, 16.475, 175.664, 3259.369, 2285.216, 42.917]
  MoveL 121 to (450, 300, 210.92) mm, rotated rx 1.89 ry 11.17 rz -178.99 deg; joints [13.984, 86.41, -173.457, -9.176, 16.032, 174.484, 3260.103, 2386.236, 43.472]
  MoveL 122 to (450, 200, 219.9) mm, rotated rx 1.62 ry 10.98 rz -179.01 deg; joints [13.984, 86.209, -173.457, -9.973, 16.397, 175.357, 3258.124, 2483.383, 51.547]
  MoveL 123 to (450, 100, 221.34) mm, rotated rx 0.64 ry 10.9 rz -179.08 deg; joints [13.984, 86.01, -173.457, -12.903, 16.632, 178.582, 3257.11, 2574.411, 51.744]
  MoveL 124 to (450, 0, 270.67) mm, rotated rx 32.3 ry 11.87 rz -176.12 deg; joints [0.856, 86.01, -173.457, 59.201, 33.971, 110.066, 3240.974, 2778.695, 176.115]
  Set speed (1000.0 mm/s)
  MoveL 125 to (450, 0, 270.67) mm, rotated rx 32.3 ry 11.87 rz -176.12 deg; joints [0.856, 86.01, -173.457, 59.201, 33.971, 110.066, 3240.974, 2778.695, 176.115]
  MoveL 126 to (470.95, -52.14, 187.95) mm, rotated rx 32.3 ry 11.87 rz -176.12 deg; joints [0.856, 86.01, -173.457, 59.201, 33.971, 110.066, 3260.969, 2831.795, 93.771]
  Set speed (1000.0 mm/s)
  MoveL 127 to (548.91, -41.08, 202.38) mm, rotated rx 25.21 ry 13.47 rz -176.13 deg; joints [3.891, 86.011, -173.457, 53.673, 27.287, 115.128, 3357.611, 2805.126, 75.591]
  MoveL 128 to (525, 0, 290.36) mm, rotated rx 25.21 ry 13.47 rz -176.13 deg; joints [3.891, 86.011, -173.457, 53.673, 27.287, 115.128, 3334.457, 2762.999, 163.279]
  MoveL 129 to (525, 0, 290.36) mm, rotated rx 25.21 ry 13.47 rz -176.13 deg; joints [3.891, 86.011, -173.457, 53.673, 27.287, 115.128, 3334.457, 2762.999, 163.279]
  Set speed (200.0 mm/s)
  MoveL 130 to (525, 100, 236.85) mm, rotated rx 0.8 ry 12.52 rz -179.04 deg; joints [13.914, 86.011, -173.457, -12.118, 15.008, 177.825, 3346.903, 2576.374, 63.83]
  MoveL 131 to (525, 200, 235.15) mm, rotated rx 1.75 ry 12.7 rz -178.95 deg; joints [13.914, 86.232, -173.457, -8.918, 14.67, 174.354, 3348.601, 2485.185, 63.447]
  MoveL 132 to (525, 300, 226.28) mm, rotated rx 2.21 ry 11.91 rz -178.94 deg; joints [13.914, 86.848, -174.321, -7.561, 15.74, 172.845, 3344.562, 2388.842, 61.889]
  MoveL 133 to (525, 400, 223.05) mm, rotated rx 1.87 ry 11.52 rz -178.98 deg; joints [14.083, 87.066, -174.626, -8.951, 16.19, 174.159, 3343.766, 2287.769, 60.885]
  MoveL 134 to (525, 500, 220.45) mm, rotated rx 1.32 ry 11.15 rz -179.03 deg; joints [14.354, 87.225, -174.85, -11.057, 16.584, 176.157, 3343.429, 2186.069, 59.85]
  MoveL 135 to (525, 600, 218.67) mm, rotated rx 0.9 ry 11.04 rz -179.06 deg; joints [14.552, 87.229, -174.85, -12.593, 16.671, 177.622, 3344.831, 2084.81, 57.555]
  MoveL 136 to (525, 700, 217.56) mm, rotated rx 0.68 ry 11 rz -179.07 deg; joints [14.658, 87.229, -174.85, -13.411, 16.7, 178.402, 3346.683, 1984.14, 55.774]
  MoveL 137 to (525, 800, 218.74) mm, rotated rx -1.55 ry 11 rz -179.23 deg; joints [15.727, 87.181, -174.782, -21.522, 16.778, 186.136, 3351.822, 1877.282, 55.774]
  MoveL 138 to (525, 900, 222) mm, rotated rx -1.77 ry 11.02 rz -179.24 deg; joints [15.823, 87.122, -174.699, -22.333, 16.753, 186.918, 3354.061, 1776.55, 57.713]
  MoveL 139 to (525, 1000, 226.01) mm, rotated rx -2.21 ry 11.97 rz -179.31 deg; joints [16.001, 86.988, -174.511, -24.429, 15.823, 188.951, 3364.872, 1674.895, 57.712]
  MoveL 140 to (525, 1100, 230.94) mm, rotated rx -2.79 ry 12.13 rz -179.37 deg; joints [16.238, 86.76, -174.191, -26.832, 15.669, 191.292, 3368.51, 1572.716, 59.455]
  MoveL 141 to (525, 1200, 236.47) mm, rotated rx -3.19 ry 12.26 rz -179.41 deg; joints [16.395, 86.595, -173.959, -28.507, 15.564, 192.93, 3371.66, 1471.164, 62.491]
  MoveL 142 to (525, 1300, 247.7) mm, rotated rx -2.64 ry 12.69 rz -179.38 deg; joints [16.395, 86.387, -173.668, -27.141, 14.968, 191.393, 3376.989, 1376.085, 69.84]
  MoveL 143 to (525, 1400, 251.45) mm, rotated rx -1.65 ry 12.56 rz -179.28 deg; joints [16.395, 86.473, -173.668, -23.827, 14.87, 187.799, 3376.99, 1284.918, 73.706]
  MoveL 144 to (525, 1500, 311.34) mm, rotated rx -22.15 ry 13.64 rz 178.22 deg; joints [23.268, 80.36, -165.33, -83.718, 24.867, 247.081, 3409.347, 1091.269, 103.416]
  Set speed (1000.0 mm/s)
  MoveL 145 to (525, 1500, 311.34) mm, rotated rx -22.15 ry 13.64 rz 178.22 deg; joints [23.268, 80.36, -165.33, -83.718, 24.867, 247.081, 3409.347, 1091.269, 103.416]
  MoveL 146 to (548, 1537.02, 221.34) mm, rotated rx -22.15 ry 13.64 rz 178.22 deg; joints [23.268, 80.36, -165.33, -83.719, 24.867, 247.081, 3433.018, 1055.316, 13.155]
  Set speed (1000.0 mm/s)
  MoveL 147 to (628.79, 1537.21, 244.37) mm, rotated rx -22.8 ry 16.82 rz 176.81 deg; joints [23.268, 78.379, -162.701, -93.295, 24.002, 256.17, 3544.956, 1051.311, 13.155]
  MoveL 148 to (600, 1500, 332.61) mm, rotated rx -22.8 ry 16.82 rz 176.81 deg; joints [23.268, 78.379, -162.701, -93.295, 24.002, 256.17, 3515.485, 1087.363, 101.652]
  MoveL 149 to (600, 1500, 332.61) mm, rotated rx -22.8 ry 16.82 rz 176.81 deg; joints [23.268, 78.379, -162.701, -93.295, 24.002, 256.17, 3515.485, 1087.363, 101.652]
  Set speed (200.0 mm/s)
  MoveL 150 to (600, 1400, 274.62) mm, rotated rx -53.63 ry 16.6 rz 168.42 deg; joints [23.268, 68.229, -149.644, -107.057, 52.228, 277.868, 3548.034, 964.026, 101.652]
  MoveL 151 to (600, 1300, 265.21) mm, rotated rx -2.11 ry 13.55 rz -179.36 deg; joints [15.353, 87.464, -175.061, -24.153, 14.305, 189.25, 3458.118, 1369.187, 96.492]
  MoveL 152 to (600, 1200, 253.06) mm, rotated rx -3.19 ry 12.8 rz -179.44 deg; joints [15.353, 87.812, -175.553, -27.137, 15.346, 192.555, 3450.308, 1459.46, 90.351]
  MoveL 153 to (600, 1100, 247.23) mm, rotated rx -3.04 ry 12.84 rz -179.42 deg; joints [15.275, 87.816, -175.559, -26.56, 15.282, 192.01, 3448.571, 1559.918, 85.14]
  MoveL 154 to (600, 1000, 242.06) mm, rotated rx -2.71 ry 13.21 rz -179.41 deg; joints [15.1, 87.816, -175.559, -25.512, 14.856, 191.031, 3449.625, 1660.776, 79.841]
  MoveL 155 to (600, 900, 237.87) mm, rotated rx -1.89 ry 13.57 rz -179.33 deg; joints [14.684, 87.816, -175.559, -22.386, 14.371, 188.079, 3449.844, 1763.078, 75.457]
  MoveL 156 to (600, 800, 234.49) mm, rotated rx -1.57 ry 11.97 rz -179.25 deg; joints [14.557, 87.816, -175.559, -20.432, 15.929, 186.188, 3432.765, 1864.372, 75.856]
  MoveL 157 to (600, 700, 233.33) mm, rotated rx 0.69 ry 11.98 rz -179.06 deg; joints [13.447, 87.864, -175.627, -11.79, 15.85, 177.982, 3427.852, 1970.986, 75.856]
  MoveL 158 to (600, 600, 234.48) mm, rotated rx 0.95 ry 12.01 rz -179.04 deg; joints [13.321, 87.864, -175.627, -10.798, 15.833, 177.039, 3425.9, 2071.723, 77.709]
  MoveL 159 to (600, 500, 236.34) mm, rotated rx 1.33 ry 12.06 rz -179.01 deg; joints [13.134, 87.864, -175.627, -9.323, 15.8, 175.638, 3424.022, 2172.825, 80.254]
  MoveL 160 to (600, 400, 239.22) mm, rotated rx 2.13 ry 12.08 rz -178.94 deg; joints [12.748, 87.864, -175.627, -6.291, 15.852, 172.755, 3421.253, 2275.163, 84.05]
  MoveL 161 to (600, 300, 242.78) mm, rotated rx 2.3 ry 12.82 rz -178.89 deg; joints [12.65, 87.584, -175.231, -5.297, 15.024, 171.826, 3425.246, 2375.681, 84.05]
  MoveL 162 to (600, 200, 252.4) mm, rotated rx 2.38 ry 13.75 rz -178.84 deg; joints [12.588, 86.947, -174.335, -4.514, 13.848, 171.106, 3430.34, 2475.951, 86.178]
  MoveL 163 to (600, 100, 254.03) mm, rotated rx 0.9 ry 13.96 rz -179.01 deg; joints [12.588, 86.797, -174.156, -10.053, 13.482, 177.062, 3430.34, 2562.923, 86.178]
  MoveL 164 to (600, 0, 311.59) mm, rotated rx 22.65 ry 15.9 rz -175.46 deg; joints [3.252, 86.797, -174.156, 57.28, 23.905, 113.435, 3432.163, 2736.265, 179.12]
  Set speed (1000.0 mm/s)
  MoveL 165 to (600, 0, 311.59) mm, rotated rx 22.65 ry 15.9 rz -175.46 deg; joints [3.252, 86.797, -174.156, 57.28, 23.905, 113.435, 3432.163, 2736.265, 179.12]
  MoveL 166 to (628.25, -36.39, 222.83) mm, rotated rx 22.65 ry 15.9 rz -175.46 deg; joints [3.252, 86.797, -174.156, 57.281, 23.905, 113.435, 3459.739, 2773.788, 90.624]
  Set speed (1000.0 mm/s)
  MoveL 167 to (712.58, -33.86, 251.33) mm, rotated rx 22.3 ry 21.19 rz -173.41 deg; joints [3.686, 84.732, -171.286, 72.055, 20.986, 99.405, 3593.386, 2773.788, 90.624]
  MoveL 168 to (675, 0, 337.6) mm, rotated rx 22.3 ry 21.19 rz -173.41 deg; joints [3.686, 84.732, -171.286, 72.055, 20.986, 99.405, 3556.436, 2738.642, 176.644]
  MoveL 169 to (675, 0, 337.6) mm, rotated rx 22.3 ry 21.19 rz -173.41 deg; joints [3.686, 84.732, -171.286, 72.055, 20.986, 99.405, 3556.436, 2738.642, 176.644]
  Set speed (200.0 mm/s)
  MoveL 170 to (675, 100, 289.19) mm, rotated rx 39.45 ry 19.85 rz -168.87 deg; joints [1.08, 84.732, -171.286, 79.758, 36.632, 90.838, 3557.37, 2738.642, 200.588]
  MoveL 171 to (675, 200, 272.28) mm, rotated rx 1.72 ry 16.92 rz -178.83 deg; joints [14.445, 85.619, -172.512, -7.866, 10.146, 172.848, 3537.533, 2494.458, 87.48]
  MoveL 172 to (675, 300, 263.14) mm, rotated rx 25.19 ry 17.48 rz -174.27 deg; joints [6.222, 84.677, -172.512, 59.363, 25.343, 108.29, 3537.533, 2494.458, 113.755]
  MoveL 173 to (675, 400, 257.86) mm, rotated rx 2.09 ry 16.04 rz -178.79 deg; joints [14.646, 84.678, -172.512, -6.397, 12, 171.061, 3541.097, 2298.24, 63.888]
  MoveL 174 to (675, 500, 254.88) mm, rotated rx 1.86 ry 14.69 rz -178.87 deg; joints [14.751, 84.844, -172.743, -8.235, 13.377, 172.829, 3530.949, 2197.341, 63.889]
  MoveL 175 to (675, 600, 253.18) mm, rotated rx 0.89 ry 14.98 rz -179 deg; joints [15.147, 84.844, -172.743, -12.404, 13.014, 176.866, 3536.758, 2093.484, 60.761]
  MoveL 176 to (675, 700, 252.08) mm, rotated rx 0.84 ry 14.94 rz -179.01 deg; joints [15.17, 84.866, -172.743, -12.676, 13.027, 177.129, 3538.133, 1993.359, 59.215]
  MoveL 177 to (675, 800, 253.29) mm, rotated rx -1.74 ry 14.93 rz -179.36 deg; joints [16.235, 84.815, -172.671, -24.182, 13.134, 188.258, 3543.375, 1883.209, 59.215]
  MoveL 178 to (675, 900, 256.88) mm, rotated rx -1.85 ry 16.51 rz -179.42 deg; joints [16.247, 84.758, -172.592, -25.821, 11.568, 189.885, 3559.914, 1782.421, 59.215]
  MoveL 179 to (675, 1000, 261.11) mm, rotated rx -2.87 ry 16.28 rz -179.58 deg; joints [16.672, 84.708, -172.523, -30.576, 11.97, 194.481, 3561.034, 1678.383, 62.826]
  MoveL 180 to (675, 1100, 266.53) mm, rotated rx -2.99 ry 16.02 rz -179.59 deg; joints [16.728, 84.708, -172.523, -30.832, 12.255, 194.719, 3560.583, 1577.965, 67.954]
  MoveL 181 to (675, 1200, 275.83) mm, rotated rx -22.66 ry 17.79 rz 176.44 deg; joints [23.548, 80.666, -167.003, -91.299, 23.442, 253.196, 3606.044, 1389.3, 67.954]
  MoveL 182 to (675, 1300, 286.17) mm, rotated rx -2.35 ry 16.54 rz -179.51 deg; joints [17.144, 82.999, -170.168, -30.734, 11.062, 194.062, 3567.724, 1389.3, 67.954]
  MoveL 183 to (675, 1400, 310.92) mm, rotated rx -32.35 ry 21.64 rz 171.85 deg; joints [23.561, 74.061, -158.292, -109.263, 31.238, 272.436, 3655.744, 1115.534, 67.954]
  Set speed (1000.0 mm/s)
  MoveL 184 to (675, 1400, 310.92) mm, rotated rx -32.35 ry 21.64 rz 171.85 deg; joints [23.561, 74.061, -158.292, -109.263, 31.238, 272.436, 3655.744, 1115.534, 67.954]
  MoveL 185 to (713.42, 1448.55, 232.39) mm, rotated rx -32.35 ry 21.64 rz 171.85 deg; joints [24.253, 75.281, -158.292, -111.772, 31.737, 274.571, 3687.267, 1081.103, 1.051]
  Set speed (1000.0 mm/s)
  MoveL 186 to (791.32, 1441.6, 268.91) mm, rotated rx -27.86 ry 23.6 rz 172.33 deg; joints [22.471, 75.281, -158.292, -114.054, 27.303, 277.175, 3772.507, 1105.567, 18.49]
  MoveL 187 to (750, 1400, 349.92) mm, rotated rx -27.86 ry 23.6 rz 172.33 deg; joints [20.4, 70.83, -158.292, -103.642, 25.698, 267.854, 3764.211, 1105.567, 57.429]
  MoveL 188 to (750, 1400, 349.92) mm, rotated rx -27.86 ry 23.6 rz 172.33 deg; joints [20.4, 70.83, -158.292, -103.642, 25.698, 267.854, 3764.211, 1105.567, 57.429]
  Set speed (200.0 mm/s)
  MoveL 189 to (750, 1300, 312.16) mm, rotated rx -2.71 ry 20.61 rz -179.76 deg; joints [16.885, 79.551, -169.871, -28.548, 9.89, 191.975, 3707.54, 1376.214, 57.429]
  MoveL 190 to (750, 1200, 303.7) mm, rotated rx -10.82 ry 20.92 rz 178.25 deg; joints [16.885, 79.551, -169.871, -62.155, 13.172, 227.09, 3709.968, 1405.79, 56.641]
  MoveL 191 to (750, 1100, 291.11) mm, rotated rx -3.1 ry 20.44 rz -179.84 deg; joints [14.642, 81.376, -172.383, -26.442, 10.742, 192.162, 3697.195, 1547.027, 56.641]
  MoveL 192 to (750, 1000, 285.42) mm, rotated rx -2.86 ry 20.75 rz -179.8 deg; joints [14.551, 81.376, -172.383, -25.502, 10.398, 191.262, 3697.99, 1648.165, 51.356]
  MoveL 193 to (750, 900, 280.81) mm, rotated rx -1.98 ry 21.15 rz -179.6 deg; joints [14.24, 81.376, -172.383, -21.065, 9.883, 186.968, 3698.994, 1752.406, 46.962]
  MoveL 194 to (750, 800, 277.21) mm, rotated rx -1.38 ry 18.58 rz -179.4 deg; joints [14.09, 81.468, -172.51, -17.056, 12.444, 183.019, 3672.53, 1855.728, 46.962]
  MoveL 195 to (750, 700, 275.91) mm, rotated rx 0.44 ry 18.58 rz -179.03 deg; joints [13.465, 81.526, -172.591, -8.804, 12.499, 175.017, 3668.988, 1964.658, 46.962]
  MoveL 196 to (750, 600, 276.71) mm, rotated rx 0.93 ry 18.76 rz -178.93 deg; joints [13.297, 81.456, -172.585, -6.493, 12.427, 172.777, 3668.988, 2066.864, 47.715]
  MoveL 197 to (750, 500, 278.49) mm, rotated rx 1.89 ry 18.63 rz -178.74 deg; joints [12.973, 81.455, -172.585, -2.328, 12.698, 168.738, 3665.03, 2171.614, 50.583]
  MoveL 198 to (750, 400, 281.44) mm, rotated rx 2.15 ry 20.48 rz -178.62 deg; joints [12.878, 81.244, -172.292, 0.767, 10.854, 165.734, 3680.133, 2272.784, 50.583]
  MoveL 199 to (750, 300, 291.13) mm, rotated rx 9.87 ry 21 rz -176.72 deg; joints [10.471, 81.243, -172.292, 33.174, 13.802, 134.358, 3678.246, 2412.156, 67.586]
  MoveL 200 to (750, 200, 296.86) mm, rotated rx 1.74 ry 20.62 rz -178.71 deg; joints [10.471, 80.549, -172.292, 1.116, 11.328, 167.876, 3678.241, 2440.362, 60.907]
  MoveL 201 to (750, 100, 327.89) mm, rotated rx 31.34 ry 23.33 rz -169.47 deg; joints [2.918, 79.231, -170.474, 74.299, 29.403, 98.188, 3704.792, 2697.231, 145.455]
  Set speed (1000.0 mm/s)
  MoveL 202 to (750, 100, 327.89) mm, rotated rx 31.34 ry 23.33 rz -169.47 deg; joints [2.918, 79.231, -170.474, 74.299, 29.403, 98.188, 3704.792, 2697.231, 145.455]
  MoveL 203 to (792.76, 55.05, 249.46) mm, rotated rx 31.34 ry 23.33 rz -169.47 deg; joints [2.918, 79.231, -170.474, 74.299, 29.403, 98.187, 3746.723, 2743.509, 67.352]
  Set speed (1000.0 mm/s)
  MoveL 204 to (875.06, 62.02, 294.05) mm, rotated rx 28.27 ry 27.97 rz -168.28 deg; joints [5.851, 76.163, -166.316, 82.951, 25.17, 87.992, 3875.398, 2741.042, 67.352]
  MoveL 205 to (825, 100, 371.84) mm, rotated rx 28.27 ry 27.97 rz -168.28 deg; joints [5.851, 76.163, -166.316, 82.951, 25.17, 87.992, 3826.037, 2701.608, 144.865]
  MoveL 206 to (825, 100, 371.84) mm, rotated rx 28.27 ry 27.97 rz -168.28 deg; joints [5.851, 76.163, -166.316, 82.951, 25.17, 87.992, 3826.037, 2701.608, 144.865]
  Set speed (200.0 mm/s)
  MoveL 207 to (825, 200, 327.16) mm, rotated rx 2.48 ry 23.88 rz -178.4 deg; joints [10.291, 78.434, -169.385, 11.215, 7.587, 157.912, 3781.731, 2446.04, 68.575]
  MoveL 208 to (825, 300, 322.5) mm, rotated rx 4.92 ry 24.58 rz -177.63 deg; joints [10.292, 78.434, -169.385, 27.797, 8.058, 140.984, 3790.367, 2367.041, 64.537]
  MoveL 209 to (825, 400, 311.37) mm, rotated rx 2.47 ry 24.85 rz -178.36 deg; joints [10.887, 79.034, -169.385, 15.039, 6.103, 153.51, 3790.387, 2253.95, 56.759]
  MoveL 210 to (825, 500, 308.31) mm, rotated rx 1.97 ry 24.92 rz -178.51 deg; joints [11.012, 79.326, -169.385, 11.823, 5.577, 156.676, 3790.424, 2151.643, 55.479]
  MoveL 211 to (825, 600, 306.59) mm, rotated rx 0.92 ry 22.95 rz -178.87 deg; joints [11.32, 79.567, -169.714, -1.525, 7.305, 169.853, 3774.482, 2046.202, 55.479]
  MoveL 212 to (825, 700, 305.89) mm, rotated rx 0.51 ry 22.75 rz -178.98 deg; joints [11.44, 79.665, -169.807, -4.742, 7.446, 173.018, 3774.482, 1944.063, 55.029]
  MoveL 213 to (825, 800, 307.3) mm, rotated rx -1.49 ry 22.73 rz -179.52 deg; joints [12.012, 79.594, -169.711, -19.257, 7.435, 187.307, 3777.558, 1833.335, 55.029]
  MoveL 214 to (825, 900, 311.14) mm, rotated rx -2.06 ry 25.2 rz -179.76 deg; joints [12.106, 79.304, -169.315, -28.871, 5.008, 196.89, 3802.825, 1729.83, 55.029]
  MoveL 215 to (825, 1000, 315.93) mm, rotated rx -2.98 ry 24.9 rz 179.96 deg; joints [12.372, 79.304, -169.315, -36.424, 5.577, 204.324, 3802.502, 1624.918, 59.358]
  MoveL 216 to (825, 1100, 322.07) mm, rotated rx -3.49 ry 24.81 rz 179.81 deg; joints [12.517, 79.285, -169.289, -40.401, 5.845, 208.237, 3803.934, 1522.16, 64.788]
  MoveL 217 to (825, 1200, 336.02) mm, rotated rx -6.42 ry 24.3 rz 178.96 deg; joints [13.358, 79.144, -169.154, -56.973, 7.787, 224.446, 3803.934, 1406.373, 78.47]
  MoveL 218 to (825, 1300, 343.92) mm, rotated rx -3.79 ry 26.61 rz 179.6 deg; joints [13.358, 78.57, -168.375, -56.934, 4.369, 223.926, 3826.812, 1329.569, 78.47]
  MoveL 219 to (825, 1400, 396.1) mm, rotated rx -32.35 ry 30.71 rz 166.68 deg; joints [15.329, 68.432, -155.051, -118.568, 28.899, 286.323, 3903.548, 1030.981, 96.942]
  Set speed (1000.0 mm/s)
  MoveL 220 to (825, 1400, 396.1) mm, rotated rx -32.35 ry 30.71 rz 166.68 deg; joints [15.329, 68.432, -155.051, -118.568, 28.899, 286.323, 3903.548, 1030.981, 96.942]
  MoveL 221 to (879.31, 1442.13, 323.47) mm, rotated rx -32.35 ry 30.71 rz 166.68 deg; joints [17.436, 73.73, -155.051, -128.002, 31.999, 294.825, 3911.486, 1030.981, 74.748]
  Set speed (1000.0 mm/s)
  MoveL 222 to (965.01, 1345.04, 338.67) mm, rotated rx -41.13 ry 35.66 rz 158.45 deg; joints [14.272, 67.774, -147.513, -134.75, 40.963, 303.605, 4063.849, 1052.925, 74.748]
  MoveL 223 to (900, 1300, 399.87) mm, rotated rx -41.13 ry 35.66 rz 158.45 deg; joints [12.661, 61.615, -147.513, -127.551, 36.751, 296.423, 4063.819, 1060.857, 78.96]
  MoveL 224 to (900, 1300, 399.87) mm, rotated rx -41.13 ry 35.66 rz 158.45 deg; joints [12.661, 61.615, -147.513, -127.551, 36.751, 296.423, 4063.819, 1060.857, 78.96]
  Set speed (200.0 mm/s)
  MoveL 225 to (900, 1200, 376.45) mm, rotated rx -5.76 ry 30.98 rz 178.53 deg; joints [12.661, 74.813, -164.49, -119.412, 4.813, 287.169, 3947.418, 1406.267, 78.96]
  MoveL 226 to (900, 1100, 361.42) mm, rotated rx -3.92 ry 32.3 rz 179.2 deg; joints [12.288, 74.813, -164.49, -143.989, 3.996, 311.895, 3956.588, 1517.577, 65.08]
  MoveL 227 to (900, 1000, 354.79) mm, rotated rx -14.05 ry 26.9 rz 157.11 deg; joints [-32.272, 78.235, -200.496, -17.821, 39, 209.606, 4213.787, 1161.862, 187.031]
  MoveL 228 to (900, 900, 349.34) mm, rotated rx -13.2 ry 27.48 rz 157.37 deg; joints [-32.375, 78.085, -200.64, -16.957, 38.461, 208.928, 4216.39, 1270.934, 180.861]
  MoveL 229 to (900, 800, 345.1) mm, rotated rx -13.01 ry 27.67 rz 157.42 deg; joints [-32.401, 78.017, -200.705, -16.771, 38.353, 208.78, 4216.459, 1373.421, 177.028]
  MoveL 230 to (900, 700, 343.45) mm, rotated rx -10.57 ry 28.58 rz 158.28 deg; joints [-32.624, 77.999, -200.723, -14.06, 36.727, 206.63, 4216.181, 1494.123, 172.897]
  MoveL 231 to (900, 600, 344.2) mm, rotated rx -9.9 ry 28.75 rz 158.52 deg; joints [-32.683, 78.04, -200.684, -13.268, 36.278, 205.994, 4213.532, 1599.163, 173.622]
  MoveL 232 to (900, 500, 346.25) mm, rotated rx 2.21 ry 29.82 rz -178.26 deg; joints [11.263, 75.247, -165.781, 62.747, 2.525, 105.588, 3924.669, 2154.676, 56.079]
  MoveL 233 to (900, 400, 349.42) mm, rotated rx 2.52 ry 29.79 rz -178.14 deg; joints [11.22, 75.019, -165.781, 59.596, 2.898, 108.755, 3924.668, 2256.231, 57.992]
  MoveL 234 to (900, 300, 360.64) mm, rotated rx 4 ry 28.77 rz -177.63 deg; joints [11.046, 73.835, -165.781, 42.791, 5.29, 125.576, 3924.668, 2364.389, 59.462]
  MoveL 235 to (900, 200, 375.7) mm, rotated rx 36.02 ry 33.05 rz -161.56 deg; joints [9.544, 70.977, -161.993, 91.85, 31.049, 77.003, 3995.671, 2681.475, 130.978]
  Set speed (1000.0 mm/s)
  MoveL 236 to (900, 200, 375.7) mm, rotated rx 36.02 ry 33.05 rz -161.56 deg; joints [9.544, 70.977, -161.993, 91.85, 31.049, 77.003, 3995.671, 2681.475, 130.978]
  MoveL 237 to (960.45, 158.17, 307.9) mm, rotated rx 36.02 ry 33.05 rz -161.56 deg; joints [9.544, 70.977, -161.993, 91.85, 31.049, 77.002, 4055.342, 2724.88, 63.491]
  Set speed (1000.0 mm/s)
  MoveL 238 to (1041.93, 291.42, 339.37) mm, rotated rx 8.94 ry 41.66 rz -173.99 deg; joints [10.264, 74.058, -161.993, 143.618, 15.526, 25.688, 4156.509, 2401.707, 63.491]
  MoveL 239 to (975, 300, 413.17) mm, rotated rx 8.94 ry 41.66 rz -173.99 deg; joints [10.264, 74.058, -161.993, 143.618, 15.526, 25.688, 4089.748, 2391.385, 137.221]
  MoveL 240 to (975, 300, 413.17) mm, rotated rx 8.94 ry 41.66 rz -173.99 deg; joints [10.264, 74.058, -161.993, 143.618, 15.526, 25.688, 4089.748, 2391.385, 137.221]
  Set speed (200.0 mm/s)
  MoveL 241 to (975, 400, 400.41) mm, rotated rx 4.06 ry 41.94 rz -176.78 deg; joints [10.774, 74.44, -161.993, 157.274, 14.713, 11.644, 4089.749, 2264.031, 124.28]
  MoveL 242 to (975, 500, 396.79) mm, rotated rx 2.59 ry 38.7 rz -177.76 deg; joints [10.961, 75.781, -163.762, 157.971, 10.9, 10.759, 4061.919, 2157.086, 124.28]
  MoveL 243 to (975, 600, 394.59) mm, rotated rx 1.93 ry 38.54 rz -178.11 deg; joints [11.066, 75.847, -163.778, 160.531, 10.693, 8.123, 4061.919, 2053.636, 121.425]
  MoveL 244 to (975, 700, 393.54) mm, rotated rx 1.21 ry 38.77 rz -178.48 deg; joints [11.162, 75.996, -163.778, 163.856, 10.995, 4.739, 4064.622, 1949.682, 121.424]
  MoveL 245 to (975, 800, 395.49) mm, rotated rx -2.48 ry 38.78 rz 179.57 deg; joints [11.767, 75.861, -163.599, 178.471, 11.194, -10.287, 4068.109, 1829.555, 121.424]
  MoveL 246 to (975, 900, 400.77) mm, rotated rx -3.18 ry 38.51 rz 179.21 deg; joints [11.898, 75.861, -163.599, 181.467, 11.062, -13.371, 4067.93, 1725.804, 125.589]
  MoveL 247 to (975, 1000, 407.69) mm, rotated rx -4.42 ry 41.61 rz 178.35 deg; joints [11.898, 74.393, -161.663, 181.713, 14.768, -13.651, 4098.624, 1618.252, 125.589]
  MoveL 248 to (975, 1100, 416.35) mm, rotated rx -5.44 ry 41.77 rz 177.76 deg; joints [12.017, 74.125, -161.311, 184.206, 15.239, -16.235, 4102.627, 1512.579, 131.886]
  MoveL 249 to (975, 1200, 433.48) mm, rotated rx -10.6 ry 42.1 rz 174.72 deg; joints [12.562, 73.019, -159.867, 195.218, 17.612, -27.654, 4111.909, 1383.404, 142.831]
  Set speed (1000.0 mm/s)
  MoveL 250 to (975, 1200, 433.48) mm, rotated rx -10.6 ry 42.1 rz 174.72 deg; joints [12.562, 73.019, -159.867, 195.218, 17.612, -27.654, 4111.909, 1383.404, 142.831]
  MoveL 251 to (1042.32, 1212.25, 360.55) mm, rotated rx -10.6 ry 42.1 rz 174.72 deg; joints [12.833, 76.294, -159.867, 192.739, 20.795, -25.317, 4147.888, 1383.404, 101.263]
  Set speed (1000.0 mm/s)
  MoveL 252 to (1072.23, 1006.4, 362.98) mm, rotated rx -5.62 ry 46.22 rz 177.3 deg; joints [11.712, 75, -158.186, 180.212, 23.524, -12.101, 4205.736, 1613.499, 101.263]
  MoveL 253 to (1000, 1000, 431.84) mm, rotated rx -5.62 ry 46.22 rz 177.3 deg; joints [11.709, 72.808, -158.186, 180.236, 21.333, -12.122, 4155.35, 1613.499, 148.926]
  MoveL 254 to (1000, 1000, 431.84) mm, rotated rx -5.62 ry 46.22 rz 177.3 deg; joints [11.709, 72.808, -158.186, 180.236, 21.333, -12.122, 4155.35, 1613.499, 148.926]
  Set speed (200.0 mm/s)
  MoveL 255 to (1000, 900, 423.58) mm, rotated rx -4.13 ry 45.18 rz 178.32 deg; joints [11.625, 73.785, -159.454, 178.162, 19.784, -9.949, 4143.083, 1721.564, 146.611]
  MoveL 256 to (1000, 800, 417.24) mm, rotated rx -2.67 ry 44.8 rz 179.23 deg; joints [11.475, 74.256, -160.068, 175.441, 19.079, -7.096, 4136.965, 1829.209, 143.845]
  MoveL 257 to (1000, 700, 414.95) mm, rotated rx 1.24 ry 44.81 rz -178.36 deg; joints [11.012, 74.428, -160.292, 167.276, 18.883, 1.449, 4133.816, 1949.479, 143.845]
  MoveL 258 to (1000, 600, 416.36) mm, rotated rx 3.06 ry 44.19 rz -177.26 deg; joints [10.845, 74.362, -160.292, 163.128, 18.314, 5.718, 4126.919, 2059.594, 143.845]
  MoveL 259 to (1000, 500, 419.51) mm, rotated rx 3.42 ry 44.95 rz -177.01 deg; joints [10.836, 73.822, -159.588, 162.817, 19.252, 6.036, 4132.099, 2161.452, 145.027]
  MoveL 260 to (1000, 400, 424.02) mm, rotated rx 5.06 ry 46.75 rz -175.87 deg; joints [10.781, 72.576, -157.971, 160.862, 21.575, 8.042, 4147.257, 2270.022, 145.129]
  Set speed (1000.0 mm/s)
  MoveL 261 to (1000, 400, 424.02) mm, rotated rx 5.06 ry 46.75 rz -175.87 deg; joints [10.781, 72.576, -157.971, 160.862, 21.575, 8.042, 4147.257, 2270.022, 145.129]
  MoveL 262 to (1073, 396.43, 355.77) mm, rotated rx 5.06 ry 46.75 rz -175.87 deg; joints [10.781, 72.574, -157.977, 160.856, 21.568, 8.048, 4220.233, 2275.392, 76.896]

--- program Top2 (robot ABB IRB 1300-10/1.15) ---
  Smooth(1)
  Set speed (1000.0 mm/s)
  Set Ref.: Top2
  Set Tool: Generic Paint Sprayer
  Show Generic Paint Sprayer
  MoveJ 1 to (1.39, -9.39, 10.94) mm, rotated rx -5.39 ry -0.83 rz -0.27 deg; joints [8.015, 137.617, -189.207, 229.616, 11.024, -53.881, 875.85, 1359.75, 0.013]
  MoveL 2 to (1.39, -9.39, 10.94) mm, rotated rx -5.39 ry -0.83 rz -0.27 deg; joints [8.015, 137.618, -189.206, 229.612, 11.025, -53.878, 875.848, 1359.75, 0.019]
  MoveL 3 to (0, 0, 110.48) mm, rotated rx -5.39 ry -0.83 rz -0.27 deg; joints [8.015, 137.618, -189.206, 229.612, 11.025, -53.878, 879.119, 1367.852, 99.635]
  MoveL 4 to (0, 0, 110.48) mm, rotated rx -5.39 ry -0.83 rz -0.27 deg; joints [8.015, 137.618, -189.206, 229.612, 11.025, -53.878, 879.119, 1367.852, 99.635]
  Set speed (200.0 mm/s)
  MoveL 5 to (0, 100, 101.49) mm, rotated rx -3.88 ry -0.62 rz -0.29 deg; joints [8.015, 137.617, -190.241, 228.699, 9.418, -53.878, 887.026, 1479.902, 86.052]
  MoveL 6 to (0, 200, 95.5) mm, rotated rx -2.82 ry -0.61 rz -0.3 deg; joints [8.015, 137.616, -190.853, 228.088, 8.275, -53.878, 890.76, 1588.523, 78.504]
  MoveL 7 to (0, 300, 91.34) mm, rotated rx -2.03 ry -0.59 rz -0.3 deg; joints [8.015, 137.616, -191.346, 227.639, 7.411, -53.878, 893.994, 1694.878, 73.418]
  MoveL 8 to (0, 400, 88.83) mm, rotated rx -1.14 ry -0.74 rz -0.3 deg; joints [8.015, 137.616, -191.723, 227.152, 6.443, -53.878, 895.014, 1802.242, 71.297]
  MoveL 9 to (0, 500, 87.56) mm, rotated rx -0.34 ry -0.73 rz -0.3 deg; joints [8.015, 137.616, -192.223, 226.708, 5.546, -53.878, 898.171, 1908.664, 69.426]
  MoveL 10 to (0, 600, 87.52) mm, rotated rx 0.56 ry -0.57 rz -0.31 deg; joints [8.015, 137.61, -192.964, 226.209, 4.501, -53.878, 904.216, 2015.674, 67.34]
  MoveL 11 to (0, 700, 89.14) mm, rotated rx 1.35 ry -0.59 rz -0.31 deg; joints [8.015, 137.409, -193.266, 225.784, 3.588, -53.878, 905.849, 2122.198, 67.339]
  MoveL 12 to (0, 800, 92.59) mm, rotated rx 2.44 ry -0.37 rz -5.31 deg; joints [6.911, 127.398, -182.498, 225.053, 5.016, -57.027, 832.992, 2205.972, 0.003]
  MoveL 13 to (0, 900, 99.11) mm, rotated rx 6.66 ry 0.27 rz -10.29 deg; joints [8.015, 134.664, -190.049, 222.478, 4.393, -61.869, 884.234, 2331.029, 62.28]
  Set speed (1000.0 mm/s)
  MoveL 14 to (0, 900, 99.11) mm, rotated rx 6.66 ry 0.27 rz -10.29 deg; joints [8.015, 134.664, -190.049, 222.478, 4.393, -61.869, 884.234, 2331.029, 62.28]
  MoveL 15 to (1.6, 911.49, -0.22) mm, rotated rx 6.66 ry 0.27 rz -10.29 deg; joints [8.015, 140.088, -195.473, 222.478, 4.393, -61.869, 920.399, 2338.225, 0.004]
  Set speed (1000.0 mm/s)
  MoveL 16 to (76.6, 911.49, 0.99) mm, rotated rx 6.66 ry 0.27 rz -10.29 deg; joints [8.015, 140.088, -195.473, 222.478, 4.393, -61.869, 845.435, 2338.191, 2.63]
  MoveL 17 to (75, 900, 100.32) mm, rotated rx 6.66 ry 0.27 rz -10.29 deg; joints [8.015, 140.088, -195.473, 222.478, 4.393, -61.869, 848.913, 2325.414, 101.749]
  MoveL 18 to (75, 900, 100.32) mm, rotated rx 6.66 ry 0.27 rz -10.29 deg; joints [8.015, 140.088, -195.473, 222.478, 4.393, -61.869, 848.913, 2325.414, 101.749]
  Set speed (200.0 mm/s)
  MoveL 19 to (75, 800, 93.37) mm, rotated rx 2.4 ry -0.4 rz -5.31 deg; joints [6.884, 129.817, -185.131, 227.279, 4.868, -59.215, 774.14, 2203.214, 20.501]
  MoveL 20 to (75, 700, 89.92) mm, rotated rx 1.4 ry -0.46 rz -5.31 deg; joints [6.884, 130.203, -184.909, 227.827, 5.99, -59.215, 772.893, 2094.818, 20.81]
  MoveL 21 to (75, 600, 88.46) mm, rotated rx 0.4 ry -0.74 rz -5.31 deg; joints [6.485, 130.203, -184.283, 228.729, 6.833, -59.215, 766.638, 1980.948, 21.319]
  MoveL 22 to (75, 500, 88.5) mm, rotated rx -0.25 ry -0.73 rz -5.3 deg; joints [6.485, 128.262, -182.035, 229.088, 7.525, -59.215, 753.086, 1877.035, 5.993]
  MoveL 23 to (75, 400, 89.77) mm, rotated rx -1.1 ry -0.81 rz -5.3 deg; joints [6.485, 128.777, -182.035, 229.499, 8.449, -59.14, 753.05, 1769.719, 12.302]
  MoveL 24 to (75, 300, 92.28) mm, rotated rx -1.73 ry -0.94 rz -5.29 deg; joints [6.485, 128.777, -181.588, 229.877, 9.142, -59.14, 749.674, 1664.489, 15.88]
  MoveL 25 to (75, 200, 96.28) mm, rotated rx -2.77 ry -0.85 rz -5.29 deg; joints [7.067, 128.789, -180.931, 229.995, 10.66, -59.14, 748.236, 1564.472, 21.154]
  MoveL 26 to (75, 100, 102.28) mm, rotated rx -2.78 ry -2.73 rz -35.25 deg; joints [8.152, 130.657, -167.078, 221.372, 36.548, -73.277, 714.805, 1372.278, 121.537]
  MoveL 27 to (75, 0, 111.64) mm, rotated rx -8.08 ry -0.98 rz -0.23 deg; joints [8.583, 130.976, -179.494, 227.194, 15.067, -50.118, 739.469, 1362.257, 70.59]
  Set speed (1000.0 mm/s)
  MoveL 28 to (75, 0, 111.64) mm, rotated rx -8.08 ry -0.98 rz -0.23 deg; joints [8.583, 130.976, -179.494, 227.194, 15.067, -50.118, 739.469, 1362.257, 70.59]
  MoveL 29 to (76.64, -14.06, 12.64) mm, rotated rx -8.08 ry -0.98 rz -0.23 deg; joints [9.696, 134.426, -182.246, 226.365, 16.085, -50.118, 757.557, 1362.257, 0]
  Set speed (1000.0 mm/s)
  MoveL 30 to (152.96, -14.2, 14.86) mm, rotated rx -8.16 ry -1.73 rz -0.12 deg; joints [9.696, 134.732, -181.692, 226.462, 16.243, -49.996, 672.011, 1362.257, 13.042]
  MoveL 31 to (150, 0, 113.8) mm, rotated rx -8.16 ry -1.73 rz -0.12 deg; joints [9.696, 134.732, -181.692, 226.462, 16.243, -49.996, 676.841, 1375.176, 112.086]
  MoveL 32 to (150, 0, 113.8) mm, rotated rx -8.16 ry -1.73 rz -0.12 deg; joints [9.696, 134.732, -181.692, 226.462, 16.243, -49.996, 676.841, 1375.176, 112.086]
  Set speed (200.0 mm/s)
  MoveL 33 to (150, 100, 104.37) mm, rotated rx -3.84 ry -1.7 rz -0.22 deg; joints [9.696, 134.732, -184.223, 223.706, 11.657, -49.996, 691.677, 1509.278, 89.224]
  MoveL 34 to (150, 200, 98.13) mm, rotated rx -2.84 ry -1.5 rz -0.25 deg; joints [9.696, 134.732, -185.087, 223.063, 10.504, -49.996, 698.429, 1616.943, 79.347]
  MoveL 35 to (150, 300, 94.12) mm, rotated rx -1.81 ry -1.47 rz -0.27 deg; joints [9.696, 134.732, -185.809, 222.44, 9.321, -49.996, 702.969, 1724.976, 73.253]
  MoveL 36 to (150, 400, 91.58) mm, rotated rx -1.16 ry -1.45 rz -0.28 deg; joints [9.696, 134.731, -186.274, 222.052, 8.56, -49.996, 705.866, 1830.05, 69.971]
  MoveL 37 to (150, 500, 90.31) mm, rotated rx -0.3 ry -1.45 rz -0.3 deg; joints [9.696, 134.731, -186.89, 221.546, 7.539, -49.996, 709.646, 1936.74, 67.489]
  MoveL 38 to (150, 600, 90.29) mm, rotated rx 0.35 ry -1.45 rz -0.31 deg; joints [9.696, 134.731, -187.36, 221.17, 6.756, -49.996, 712.496, 2041.781, 66.995]
  MoveL 39 to (150, 700, 91.77) mm, rotated rx 1.38 ry -1.47 rz -0.33 deg; joints [9.696, 134.711, -188.096, 220.581, 5.494, -49.996, 716.92, 2149.769, 66.994]
  MoveL 40 to (150, 800, 95.46) mm, rotated rx 2.37 ry -1.67 rz -0.36 deg; joints [9.163, 134.313, -188.592, 220.472, 3.832, -49.996, 716.92, 2250.424, 66.995]
  MoveL 41 to (150, 900, 102.49) mm, rotated rx 6.81 ry -1.08 rz -5.42 deg; joints [13.295, 132.635, -185.769, 220.549, 5.415, -60.054, 710.315, 2426.711, 68.287]
  Set speed (1000.0 mm/s)
  MoveL 42 to (150, 900, 102.49) mm, rotated rx 6.81 ry -1.08 rz -5.42 deg; joints [13.295, 132.635, -185.769, 220.549, 5.415, -60.054, 710.315, 2426.711, 68.287]
  MoveL 43 to (152.99, 911.63, 3.22) mm, rotated rx 6.81 ry -1.08 rz -5.42 deg; joints [13.295, 136.955, -190.089, 220.549, 5.415, -60.054, 735.169, 2432.607, 0]
  Set speed (1000.0 mm/s)
  MoveL 44 to (229.53, 911.76, 6.23) mm, rotated rx 6.98 ry -1.95 rz -5.52 deg; joints [13.187, 137.113, -189.26, 220.62, 5.568, -60.054, 646.044, 2432.607, 13.361]
  MoveL 45 to (225, 900, 105.43) mm, rotated rx 6.98 ry -1.95 rz -5.52 deg; joints [13.187, 137.113, -189.26, 220.619, 5.568, -60.054, 652.446, 2419.56, 112.299]
  MoveL 46 to (225, 900, 105.43) mm, rotated rx 6.98 ry -1.95 rz -5.52 deg; joints [13.187, 137.113, -189.26, 220.619, 5.568, -60.054, 652.446, 2419.56, 112.299]
  Set speed (200.0 mm/s)
  MoveL 47 to (225, 800, 98.09) mm, rotated rx 2.61 ry -2.26 rz -0.39 deg; joints [9.088, 142.739, -196.781, 222.709, 3.449, -52.283, 697.877, 2241.517, 130.6]
  MoveL 48 to (225, 700, 94.38) mm, rotated rx 1.38 ry -2.37 rz -0.35 deg; joints [9.088, 143.638, -196.694, 223.407, 4.926, -52.283, 697.875, 2131.039, 134.775]
  MoveL 49 to (225, 600, 92.87) mm, rotated rx 0.35 ry -2.34 rz -0.32 deg; joints [9.088, 144.125, -196.517, 223.999, 6.116, -52.283, 697.874, 2022.38, 137.086]
  MoveL 50 to (225, 500, 92.76) mm, rotated rx -0.3 ry -2.19 rz -0.3 deg; joints [9.088, 144.163, -196.299, 224.365, 6.831, -52.283, 697.874, 1917.097, 136.196]
  MoveL 51 to (225, 400, 94.03) mm, rotated rx -1.16 ry -2.2 rz -0.27 deg; joints [9.088, 144.584, -196.166, 224.872, 7.801, -52.283, 697.872, 1809.812, 140.877]
  MoveL 52 to (225, 300, 96.7) mm, rotated rx -1.81 ry -2.36 rz -0.24 deg; joints [9.088, 145.162, -196.166, 225.276, 8.547, -52.283, 697.758, 1704.116, 148.73]
  MoveL 53 to (225, 200, 100.75) mm, rotated rx -2.84 ry -2.39 rz -0.21 deg; joints [9.088, 145.68, -196.024, 225.901, 9.673, -52.283, 697.757, 1595.37, 157.59]
  MoveL 54 to (225, 100, 106.98) mm, rotated rx -4.07 ry -2.3 rz -0.17 deg; joints [9.088, 146.011, -195.746, 226.644, 10.979, -52.283, 697.755, 1485.017, 167.046]
  MoveL 55 to (225, 0, 116.73) mm, rotated rx -8.27 ry -2.63 rz 0.01 deg; joints [9.088, 148.107, -195.313, 229.367, 15.274, -52.283, 697.753, 1349.343, 202.943]
  Set speed (1000.0 mm/s)
  MoveL 56 to (225, 0, 116.73) mm, rotated rx -8.27 ry -2.63 rz 0.01 deg; joints [9.088, 148.107, -195.313, 229.367, 15.274, -52.283, 697.753, 1349.343, 202.943]
  MoveL 57 to (229.54, -14.38, 17.88) mm, rotated rx -8.27 ry -2.63 rz 0.01 deg; joints [9.088, 148.107, -195.313, 229.367, 15.274, -52.283, 691.349, 1336.239, 104.013]
  Set speed (1000.0 mm/s)
  MoveL 58 to (306.2, -14.36, 21.68) mm, rotated rx -8.27 ry -3.57 rz 0.15 deg; joints [9.075, 149.053, -195.313, 229.568, 15.289, -52.283, 609.328, 1336.24, 122.863]
  MoveL 59 to (300, 0, 120.45) mm, rotated rx -8.27 ry -3.57 rz 0.15 deg; joints [9.075, 149.053, -195.313, 229.568, 15.289, -52.283, 617.395, 1349.321, 221.674]
  MoveL 60 to (300, 0, 120.45) mm, rotated rx -8.27 ry -3.57 rz 0.15 deg; joints [9.075, 149.053, -195.313, 229.568, 15.289, -52.283, 617.395, 1349.321, 221.674]
  Set speed (200.0 mm/s)
  MoveL 61 to (300, 100, 110.26) mm, rotated rx -3.88 ry -3.2 rz -0.12 deg; joints [9.075, 146.876, -195.766, 226.669, 10.875, -52.283, 617.396, 1486.252, 184.131]
  MoveL 62 to (300, 200, 104.08) mm, rotated rx -2.85 ry -3.14 rz -0.17 deg; joints [9.075, 146.379, -195.909, 226.02, 9.783, -52.283, 617.396, 1594.975, 173.096]
  MoveL 63 to (300, 300, 99.81) mm, rotated rx -1.96 ry -2.97 rz -0.22 deg; joints [9.075, 145.695, -195.937, 225.452, 8.802, -52.283, 617.396, 1702.677, 162.265]
  MoveL 64 to (300, 400, 97.17) mm, rotated rx -1.16 ry -3.09 rz -0.25 deg; joints [9.075, 145.555, -196.158, 224.977, 7.941, -52.283, 617.396, 1809.291, 159.044]
  MoveL 65 to (300, 500, 95.9) mm, rotated rx -0.29 ry -3.08 rz -0.29 deg; joints [9.075, 145.147, -196.298, 224.455, 6.978, -52.283, 617.396, 1916.581, 154.448]
  MoveL 66 to (300, 600, 95.99) mm, rotated rx 0.51 ry -2.96 rz -0.33 deg; joints [9.075, 144.529, -196.335, 223.97, 6.051, -52.283, 617.397, 2023.456, 149.155]
  MoveL 67 to (300, 700, 97.71) mm, rotated rx 1.41 ry -3.12 rz -0.37 deg; joints [9.075, 144.375, -196.597, 223.455, 5.053, -52.283, 617.397, 2130.742, 150.554]
  MoveL 68 to (300, 800, 101.35) mm, rotated rx 2.43 ry -3.16 rz -0.42 deg; joints [9.075, 143.909, -196.784, 222.868, 3.87, -52.283, 617.396, 2239.189, 150.758]
  MoveL 69 to (300, 900, 109.13) mm, rotated rx 7.46 ry -1.65 rz -15.57 deg; joints [10.775, 142.611, -191.132, 219.696, 11.224, -65.537, 589.136, 2344.943, 166.949]
  Set speed (1000.0 mm/s)
  MoveL 70 to (300, 900, 109.13) mm, rotated rx 7.06 ry -2.91 rz -5.64 deg; joints [12.922, 124.127, -174.581, 216.956, 6.21, -56.124, 475.851, 2436.699, 30.038]
  MoveL 71 to (306.23, 911.74, 10.02) mm, rotated rx 7.06 ry -2.91 rz -5.64 deg; joints [12.922, 132.894, -183.348, 216.956, 6.21, -56.124, 521.096, 2437.484, 0.001]
  Set speed (1000.0 mm/s)
  MoveL 72 to (381.1, 911.97, 14.67) mm, rotated rx 7.19 ry -2.83 rz -5.64 deg; joints [12.922, 132.894, -183.55, 216.874, 6.008, -56.124, 448.135, 2438.511, 4.989]
  MoveL 73 to (375, 900, 113.76) mm, rotated rx 7.19 ry -2.83 rz -5.64 deg; joints [12.922, 132.894, -183.549, 216.874, 6.008, -56.124, 456.107, 2425.256, 103.785]
  MoveL 74 to (375, 900, 113.76) mm, rotated rx 7.19 ry -2.83 rz -5.64 deg; joints [12.922, 132.894, -183.549, 216.874, 6.008, -56.124, 456.107, 2425.256, 103.785]
  Set speed (200.0 mm/s)
  MoveL 75 to (375, 800, 105.52) mm, rotated rx 2.43 ry -3.16 rz -0.42 deg; joints [9, 143.644, -196.792, 225.326, 3.643, -54.687, 541.937, 2238.261, 153.707]
  MoveL 76 to (375, 700, 101.74) mm, rotated rx 1.59 ry -2.98 rz -0.37 deg; joints [9.014, 143.701, -196.528, 225.786, 4.561, -54.687, 541.937, 2131.713, 149.017]
  MoveL 77 to (375, 600, 99.96) mm, rotated rx 0.38 ry -3.09 rz -0.32 deg; joints [9.014, 144.474, -196.448, 226.497, 5.921, -54.687, 541.937, 2021.415, 154.089]
  MoveL 78 to (375, 500, 99.93) mm, rotated rx -0.29 ry -3.08 rz -0.29 deg; joints [9.013, 144.753, -196.348, 226.887, 6.639, -54.687, 541.936, 1915.861, 155.795]
  MoveL 79 to (375, 400, 101.2) mm, rotated rx -1.16 ry -3.08 rz -0.25 deg; joints [9.013, 145.131, -196.223, 227.409, 7.58, -54.687, 541.935, 1808.496, 160.025]
  MoveL 80 to (375, 300, 103.79) mm, rotated rx -1.83 ry -3.1 rz -0.22 deg; joints [9.013, 145.422, -196.133, 227.806, 8.284, -54.684, 541.933, 1702.9, 164.705]
  MoveL 81 to (375, 200, 108.1) mm, rotated rx -3.04 ry -2.99 rz -0.17 deg; joints [9.013, 145.7, -195.875, 228.53, 9.533, -54.684, 541.932, 1592.825, 171.371]
  MoveL 82 to (375, 100, 114.43) mm, rotated rx -3.88 ry -3.2 rz -0.12 deg; joints [9.014, 146.35, -195.875, 229.075, 10.42, -54.684, 541.821, 1485.524, 184.082]
  MoveL 83 to (375, 0, 125.12) mm, rotated rx -8.33 ry -3.54 rz 0.15 deg; joints [9.03, 148.85, -195.254, 229.95, 15.239, -52.608, 541.817, 1348.263, 225.949]
  Set speed (1000.0 mm/s)
  MoveL 84 to (375, 0, 125.12) mm, rotated rx -8.33 ry -3.54 rz 0.15 deg; joints [9.03, 148.85, -195.254, 229.95, 15.239, -52.608, 541.817, 1348.263, 225.949]
  MoveL 85 to (381.14, -14.47, 26.36) mm, rotated rx -8.33 ry -3.54 rz 0.15 deg; joints [9.03, 148.85, -195.254, 229.95, 15.239, -52.608, 533.812, 1335.067, 127.148]
  Set speed (1000.0 mm/s)
  MoveL 86 to (457.45, -14.94, 32.13) mm, rotated rx -8.62 ry -4.28 rz 0.28 deg; joints [9.03, 149.833, -195.254, 230, 15.593, -52.304, 454.167, 1332.215, 147.781]
  MoveL 87 to (450, 0, 130.73) mm, rotated rx -8.04 ry 5.28 rz 59.58 deg; joints [23.35, 135.017, -168.997, 162.83, 31.392, 51.519, 460.58, 1780.09, 178.693]
  MoveL 88 to (450, 0, 130.73) mm, rotated rx -8.95 ry -3.52 rz 5.23 deg; joints [-0.797, 145.171, -196.599, 229.742, 4.914, -40.555, 452.096, 1244.299, 192.082]
  Set speed (200.0 mm/s)
  MoveL 89 to (450, 100, 119.63) mm, rotated rx -5.49 ry 1.34 rz 59.74 deg; joints [23.35, 135.188, -168.476, 154.815, 31.392, 56.695, 460.58, 1921.939, 185.652]
  MoveL 90 to (450, 200, 113.07) mm, rotated rx -2.89 ry -4.02 rz -0.12 deg; joints [-12.753, 136.541, -196.259, 50, 7.007, 141.577, 457.839, 1321.957, 89.663]
  MoveL 91 to (450, 300, 108.84) mm, rotated rx -1.98 ry -3.85 rz -0.19 deg; joints [-12.753, 135.76, -196.395, 50, 7.939, 141.167, 459.636, 1429.695, 77.469]
  MoveL 92 to (450, 400, 106.11) mm, rotated rx -1.17 ry -3.84 rz -0.24 deg; joints [-12.753, 138.859, -200.203, 50, 8.806, 140.8, 486.725, 1542.597, 94.805]
  MoveL 93 to (450, 500, 104.84) mm, rotated rx -0.28 ry -3.83 rz -0.29 deg; joints [-12.753, 138.168, -200.273, 49.999, 9.759, 140.407, 486.726, 1650.003, 88.016]
  MoveL 94 to (450, 600, 105.02) mm, rotated rx 0.53 ry -3.84 rz -0.34 deg; joints [-13, 143.068, -206.005, 50, 10.82, 140.276, 529.918, 1763.675, 118.478]
  MoveL 95 to (450, 700, 106.7) mm, rotated rx 1.59 ry -3.88 rz -0.4 deg; joints [-6.6, 149.984, -210, 50, 7.231, 134.101, 554.728, 1948.633, 168.758]
  MoveL 96 to (450, 800, 110.76) mm, rotated rx 4.04 ry -4.45 rz 4.41 deg; joints [-0.797, 139.286, -200.351, 48.296, 9.468, 133.954, 469.454, 2152.632, 113.1]
  MoveL 97 to (450, 900, 119.35) mm, rotated rx 7.17 ry -4.21 rz -0.78 deg; joints [7.013, 154.124, -210, 50, 2.958, 119.654, 561.525, 2339.246, 223.094]
  Set speed (1000.0 mm/s)
  MoveL 98 to (450, 900, 119.35) mm, rotated rx 7.17 ry -4.21 rz -0.78 deg; joints [7.013, 154.124, -210, 50, 2.958, 119.654, 561.525, 2339.246, 223.094]
  MoveL 99 to (457.45, 912.39, 20.4) mm, rotated rx 7.17 ry -4.21 rz -0.78 deg; joints [7.013, 143.846, -199.722, 50, 2.958, 119.654, 464.59, 2363.694, 71.395]
  Set speed (1000.0 mm/s)
  MoveL 100 to (534.03, 912.36, 26.81) mm, rotated rx 6.71 ry -5.72 rz 4.09 deg; joints [-0.912, 138.714, -200.634, 48.282, 12.552, 132.684, 376.794, 2286.663, 34.465]
  MoveL 101 to (525, 900, 125.63) mm, rotated rx 6.71 ry -5.72 rz 4.09 deg; joints [-0.912, 138.714, -200.634, 48.282, 12.552, 132.684, 387.689, 2273.024, 132.929]
  MoveL 102 to (525, 900, 125.63) mm, rotated rx 6.71 ry -5.72 rz 4.09 deg; joints [-0.912, 138.714, -200.634, 48.282, 12.552, 132.684, 387.689, 2273.024, 132.929]
  Set speed (200.0 mm/s)
  MoveL 103 to (525, 800, 116.73) mm, rotated rx 4.02 ry -5.23 rz 4.36 deg; joints [-0.388, 140.143, -200.172, 48.282, 9.152, 133.52, 387.689, 2157.531, 132.929]
  MoveL 104 to (525, 700, 112.5) mm, rotated rx 1.04 ry -4.88 rz 4.6 deg; joints [-0.439, 141.708, -199.801, 48.313, 5.877, 135.021, 387.689, 2032.385, 140.417]
  MoveL 105 to (525, 600, 110.59) mm, rotated rx 0.13 ry -4.62 rz 4.67 deg; joints [0.123, 141.558, -198.863, 48.313, 4.421, 135.021, 382.708, 1931.697, 137.531]
  MoveL 106 to (525, 500, 110.39) mm, rotated rx -0.67 ry -4.54 rz 4.73 deg; joints [0.123, 141.566, -198.318, 48.346, 3.521, 135.411, 379.288, 1825.016, 137.531]
  MoveL 107 to (525, 400, 111.66) mm, rotated rx -1.56 ry -4.46 rz 4.79 deg; joints [0.117, 142.086, -198.209, 48.371, 2.543, 135.861, 379.288, 1717.592, 142.661]
  MoveL 108 to (525, 300, 114.42) mm, rotated rx -4.01 ry -3 rz 29.86 deg; joints [39.036, 151.866, -200.177, -133.306, 11.749, 308.211, 591.49, 2127.558, 223.73]
  MoveL 109 to (525, 200, 118.88) mm, rotated rx -2.89 ry -4.79 rz -0.09 deg; joints [14.34, 134.152, -180.793, -130, 13.438, 299.958, 284.456, 1686.495, 134.426]
  MoveL 110 to (525, 100, 125.58) mm, rotated rx -5.9 ry -4.91 rz 0.16 deg; joints [17.159, 134.154, -178.049, -130, 18.798, 299.958, 279.583, 1605.466, 155.048]
  MoveL 111 to (525, 0, 137.03) mm, rotated rx -8.9 ry -5.03 rz 0.41 deg; joints [20.263, 134.155, -175.288, -130.015, 24.387, 299.958, 279.065, 1529.28, 182.583]
  Set speed (1000.0 mm/s)
  MoveL 112 to (525, 0, 137.03) mm, rotated rx -8.9 ry -5.03 rz 0.41 deg; joints [20.263, 134.155, -175.288, -130.015, 24.387, 299.958, 279.065, 1529.28, 182.583]
  MoveL 113 to (533.77, -15.42, 38.62) mm, rotated rx -8.9 ry -5.03 rz 0.41 deg; joints [20.263, 134.155, -175.288, -130.015, 24.387, 299.958, 268.434, 1515.139, 84.161]
  Set speed (1000.0 mm/s)
  MoveL 114 to (610.79, -15.37, 45.77) mm, rotated rx -8.91 ry -6.18 rz 0.59 deg; joints [20.175, 135.03, -174.765, -130, 24.639, 300.449, 180.513, 1515.139, 111.95]
  MoveL 115 to (600, 0, 143.99) mm, rotated rx -8.91 ry -6.18 rz 0.59 deg; joints [20.17, 135.03, -174.761, -130.009, 24.639, 300.463, 193.111, 1529.179, 210.163]
  MoveL 116 to (600, 0, 143.99) mm, rotated rx -8.91 ry -6.18 rz 0.59 deg; joints [20.17, 135.03, -174.761, -130.009, 24.639, 300.463, 193.111, 1529.179, 210.163]
  Set speed (200.0 mm/s)
  MoveL 117 to (600, 100, 132.29) mm, rotated rx -6.19 ry -5.81 rz 0.28 deg; joints [20.17, 135.03, -175.712, -132.033, 22.331, 300.463, 200.742, 1649.251, 190.183]
  MoveL 118 to (600, 200, 125.29) mm, rotated rx -3.1 ry -5.69 rz -0.02 deg; joints [20.17, 135.03, -176.625, -134.193, 19.618, 300.463, 206.209, 1772.724, 177.389]
  MoveL 119 to (600, 300, 120.71) mm, rotated rx -1.98 ry -5.66 rz -0.12 deg; joints [20.17, 135.03, -176.981, -134.958, 18.604, 300.463, 208.181, 1881.2, 171.838]
  MoveL 120 to (600, 400, 118.12) mm, rotated rx -0.92 ry -5.48 rz -0.22 deg; joints [20.17, 135.03, -177.515, -135.722, 17.568, 300.463, 212.283, 1988.912, 166.874]
  MoveL 121 to (600, 500, 116.83) mm, rotated rx -0.51 ry -5.48 rz -0.26 deg; joints [20.17, 135.03, -177.647, -135.993, 17.191, 300.463, 212.951, 2091.963, 166.211]
  MoveL 122 to (600, 600, 116.88) mm, rotated rx 0.55 ry -5.64 rz -0.35 deg; joints [20.17, 135.03, -177.803, -136.663, 16.245, 300.463, 212.362, 2200.355, 167.719]
  MoveL 123 to (600, 700, 118.91) mm, rotated rx 1.67 ry -5.66 rz -0.46 deg; joints [20.17, 134.769, -177.916, -137.4, 15.18, 300.463, 212.436, 2309.34, 167.719]
  MoveL 124 to (600, 800, 123.43) mm, rotated rx 4.74 ry -5.76 rz -0.75 deg; joints [20.17, 134.374, -178.6, -139.392, 12.164, 300.463, 214.592, 2433.104, 167.719]
  MoveL 125 to (600, 900, 132.59) mm, rotated rx 7.44 ry -6.13 rz -1.05 deg; joints [20.17, 134.263, -179.202, -141.066, 9.532, 300.463, 214.592, 2553.373, 178.535]
  Set speed (1000.0 mm/s)
  MoveL 126 to (600, 900, 132.59) mm, rotated rx 7.44 ry -6.13 rz -1.05 deg; joints [20.17, 134.263, -179.202, -141.066, 9.532, 300.463, 214.592, 2553.373, 178.535]
  MoveL 127 to (610.82, 912.76, 34) mm, rotated rx 7.44 ry -6.13 rz -1.05 deg; joints [20.17, 134.263, -179.202, -141.066, 9.532, 300.463, 201.915, 2567.407, 80.339]
  Set speed (1000.0 mm/s)
  MoveL 128 to (685.68, 913.03, 42.2) mm, rotated rx 7.6 ry -6.04 rz -1.05 deg; joints [20.17, 134.263, -179.388, -141.177, 9.319, 300.462, 128.866, 2568.503, 88.852]
  MoveL 129 to (675, 900, 140.77) mm, rotated rx 7.6 ry -6.04 rz -1.05 deg; joints [20.17, 134.263, -179.388, -141.177, 9.319, 300.462, 141.404, 2554.198, 187.026]
  MoveL 130 to (675, 900, 140.77) mm, rotated rx 7.6 ry -6.04 rz -1.05 deg; joints [20.17, 134.263, -179.388, -141.177, 9.319, 300.462, 141.404, 2554.198, 187.026]
  Set speed (200.0 mm/s)
  MoveL 131 to (675, 800, 131.08) mm, rotated rx 4.74 ry -5.76 rz -0.75 deg; joints [20.17, 134.624, -178.851, -139.391, 12.163, 300.462, 141.404, 2432.378, 178.566]
  MoveL 132 to (675, 700, 126.36) mm, rotated rx 1.67 ry -5.66 rz -0.46 deg; joints [20.17, 135.05, -178.2, -137.4, 15.179, 300.462, 139.478, 2308.544, 178.566]
  MoveL 133 to (675, 600, 124.2) mm, rotated rx 0.73 ry -5.48 rz -0.37 deg; joints [20.17, 135.05, -178.084, -136.821, 16.012, 300.462, 140.319, 2201.194, 174.537]
  MoveL 134 to (675, 500, 124.02) mm, rotated rx -0.51 ry -5.47 rz -0.26 deg; joints [20.17, 135.05, -177.671, -135.994, 17.188, 300.462, 138.27, 2091.813, 174.925]
  MoveL 135 to (675, 400, 125.31) mm, rotated rx -0.92 ry -5.48 rz -0.22 deg; joints [20.17, 135.05, -177.538, -135.72, 17.569, 300.462, 137.601, 1988.723, 175.592]
  MoveL 136 to (675, 300, 128.03) mm, rotated rx -2.16 ry -5.5 rz -0.11 deg; joints [20.17, 135.05, -177.131, -134.881, 18.717, 300.462, 135.418, 1879.326, 179.318]
  MoveL 137 to (675, 200, 132.76) mm, rotated rx -3.11 ry -5.68 rz -0.02 deg; joints [20.17, 135.051, -176.651, -134.188, 19.623, 300.462, 131.582, 1772.475, 186.35]
  MoveL 138 to (675, 100, 139.96) mm, rotated rx -6.19 ry -5.81 rz 0.28 deg; joints [20.17, 135.051, -175.733, -132.032, 22.331, 300.462, 126.037, 1649.083, 199.402]
  MoveL 139 to (675, 0, 152.2) mm, rotated rx -8.99 ry -6.14 rz 0.59 deg; joints [20.223, 135.051, -174.775, -130, 24.75, 300.462, 118.986, 1529.082, 219.854]
  Set speed (1000.0 mm/s)
  MoveL 140 to (675, 0, 152.2) mm, rotated rx -8.99 ry -6.14 rz 0.59 deg; joints [20.223, 135.051, -174.775, -130, 24.75, 300.462, 118.986, 1529.082, 219.854]
  MoveL 141 to (685.72, -15.51, 54) mm, rotated rx -8.99 ry -6.14 rz 0.59 deg; joints [20.223, 135.051, -174.775, -130, 24.75, 300.462, 106.414, 1514.844, 121.675]
  Set speed (1000.0 mm/s)
  MoveL 142 to (761.71, -16.08, 63.23) mm, rotated rx -9.34 ry -6.7 rz 0.72 deg; joints [20.384, 135.472, -174.237, -130, 25.407, 300.849, 24.97, 1514.714, 143.678]
  MoveL 143 to (750, 0, 161.23) mm, rotated rx -9.34 ry -6.7 rz 0.72 deg; joints [-4.974, 135.472, -183.618, -130, 5.192, 318.858, 40.303, 1160.164, 195.683]
  MoveL 144 to (750, 0, 161.23) mm, rotated rx -9.34 ry -6.7 rz 0.72 deg; joints [-4.974, 135.472, -183.618, -130, 5.192, 318.858, 40.303, 1160.164, 195.683]
  Set speed (200.0 mm/s)
  MoveL 145 to (750, 100, 148.42) mm, rotated rx -6.9 ry -5.9 rz 5.36 deg; joints [-0.682, 153.628, -204.163, -137.614, 2.666, 325.535, 202.013, 1365.942, 272.818]
  MoveL 146 to (750, 200, 140.94) mm, rotated rx -2.54 ry -6.57 rz -5.01 deg; joints [13.221, 136.756, -177.555, -136.348, 18.258, 303.874, 30.793, 1652.541, 215.864]
  MoveL 147 to (750, 300, 136.06) mm, rotated rx -1.62 ry -6.37 rz -5.11 deg; joints [13.221, 136.756, -178.12, -137.033, 17.348, 303.874, 34.597, 1759.404, 208.204]
  MoveL 148 to (750, 400, 133.14) mm, rotated rx -0.67 ry -5.93 rz -5.22 deg; joints [13.221, 136.756, -179.008, -137.792, 16.304, 303.874, 42.09, 1866.315, 199.832]
  MoveL 149 to (750, 500, 131.86) mm, rotated rx 0.27 ry -5.84 rz -5.31 deg; joints [13.221, 136.756, -179.504, -138.451, 15.349, 303.874, 44.725, 1973.412, 197.024]
  MoveL 150 to (750, 600, 132.23) mm, rotated rx 1.29 ry -6.11 rz -5.41 deg; joints [13.221, 136.756, -179.626, -139.079, 14.426, 303.874, 42.512, 2081.245, 199.629]
  MoveL 151 to (750, 700, 134.54) mm, rotated rx 2.22 ry -6.13 rz -5.5 deg; joints [13.221, 136.581, -179.839, -139.698, 13.493, 303.874, 42.511, 2188.471, 200.591]
  MoveL 152 to (750, 800, 139.52) mm, rotated rx 5.47 ry -5.98 rz -5.83 deg; joints [13.221, 136.581, -181.656, -141.873, 9.988, 303.874, 51.318, 2312.293, 199.553]
  MoveL 153 to (750, 900, 149.76) mm, rotated rx 8.17 ry -6.12 rz -6.14 deg; joints [13.221, 135.959, -182.375, -143.596, 7.019, 303.874, 51.318, 2432.687, 204.287]
  Set speed (1000.0 mm/s)
  MoveL 154 to (750, 900, 149.76) mm, rotated rx 8.17 ry -6.12 rz -6.14 deg; joints [13.221, 135.959, -182.375, -143.596, 7.019, 303.874, 51.318, 2432.687, 204.287]
  MoveL 155 to (762.02, 913, 51.34) mm, rotated rx 8.17 ry -6.12 rz -6.14 deg; joints [13.221, 135.959, -182.375, -143.596, 7.019, 303.874, 37.446, 2446.953, 106.287]

--- program DoorRR_C (robot ABB IRB 1300-10/1.15) ---
  Smooth(1)
  Set speed (1000.0 mm/s)
  Set Ref.: DoorRR
  Set Tool: Generic Paint Sprayer
  Show Generic Paint Sprayer
  MoveJ 1 to (-63.47, 907.08, 255.99) mm, rotated rx 39.6 ry -2.99 rz 87.24 deg; joints [-128.12, 34.671, -33.35, 123.573, 79.803, -211.755, 1679.755, -179.592, 100.569]
  MoveL 2 to (-63.47, 907.08, 255.99) mm, rotated rx 39.6 ry -2.99 rz 87.24 deg; joints [-128.12, 34.671, -33.35, 123.573, 79.803, -211.755, 1679.757, -179.593, 100.574]
  MoveL 3 to (0, 900, 332.94) mm, rotated rx 39.6 ry -2.99 rz 87.24 deg; joints [-127.915, 34.535, -33.35, 123.577, 79.558, -211.755, 1679.759, -103.507, 162.351]
  MoveL 4 to (0, 900, 332.94) mm, rotated rx 39.6 ry -2.99 rz 87.24 deg; joints [-127.915, 34.535, -33.35, 123.577, 79.558, -211.755, 1679.759, -103.507, 162.351]
  Set speed (200.0 mm/s)
  MoveL 5 to (0, 800, 323.94) mm, rotated rx 38.28 ry -2.84 rz 87.41 deg; joints [-127.915, 34.519, -33.35, 122.717, 78.783, -210.888, 1781.675, -117.398, 172.973]
  MoveL 6 to (0, 700, 315.56) mm, rotated rx 37.73 ry -2.69 rz 87.55 deg; joints [-127.915, 34.519, -33.35, 122.423, 78.367, -210.547, 1883.605, -126.592, 178.774]
  MoveL 7 to (0, 600, 307.63) mm, rotated rx 36.98 ry -2.66 rz 87.59 deg; joints [-127.915, 34.516, -33.35, 121.882, 78.004, -210.043, 1984.114, -135.826, 186.427]
  MoveL 8 to (0, 500, 300.04) mm, rotated rx 32.16 ry -2.81 rz 87.64 deg; joints [-127.915, 34.515, -33.133, 118.177, 76.235, -206.887, 2083.534, -163.643, 224.679]
  MoveL 9 to (0, 400, 292.72) mm, rotated rx 31.37 ry -2.7 rz 87.73 deg; joints [-127.915, 34.515, -33.133, 117.621, 75.809, -206.341, 2184.841, -172.291, 232.801]
  MoveL 10 to (0, 300, 285.76) mm, rotated rx 30.76 ry -2.51 rz 87.86 deg; joints [-127.915, 34.515, -33.133, 117.245, 75.373, -205.932, 2286.918, -180.036, 239.468]
  MoveL 11 to (0, 200, 279.5) mm, rotated rx 29.26 ry -2.34 rz 87.99 deg; joints [-127.915, 34.515, -33.133, 116.14, 74.636, -204.876, 2388.784, -190.713, 252.814]
  MoveL 12 to (0, 100, 273.72) mm, rotated rx 28.63 ry -2.21 rz 88.07 deg; joints [-127.915, 34.515, -33.133, 115.701, 74.269, -204.437, 2490.209, -196.947, 259.916]
  MoveL 13 to (0, 0, 268.4) mm, rotated rx 25.03 ry -2.21 rz 88.12 deg; joints [-127.915, 34.514, -33.133, 112.751, 73.035, -201.769, 2590.477, -213.484, 290.009]
  Set speed (1000.0 mm/s)
  MoveL 14 to (0, 0, 268.4) mm, rotated rx 25.03 ry -2.21 rz 88.12 deg; joints [-127.915, 34.514, -33.133, 112.751, 73.035, -201.769, 2590.477, -213.484, 290.009]
  MoveL 15 to (-42.18, 4.87, 177.86) mm, rotated rx 25.03 ry -2.21 rz 88.12 deg; joints [-128.003, 34.551, -33.133, 112.748, 73.13, -201.769, 2590.477, -303.537, 248.292]
  Set speed (1000.0 mm/s)
  MoveL 16 to (77.33, 5.4, 118.5) mm, rotated rx -1.25 ry -3.13 rz 88.47 deg; joints [-131.414, 29.408, -33.133, 87.7, 73.13, -175.081, 2590.477, -334.567, 520.202]
  MoveL 17 to (75, 0, 218.33) mm, rotated rx -1.25 ry -3.13 rz 88.47 deg; joints [-131.159, 29.418, -33.133, 87.684, 72.876, -175.081, 2590.478, -237.209, 518.043]
  MoveL 18 to (75, 0, 218.33) mm, rotated rx -1.25 ry -3.13 rz 88.47 deg; joints [-131.159, 29.418, -33.133, 87.684, 72.876, -175.081, 2590.478, -237.209, 518.043]
  Set speed (200.0 mm/s)
  MoveL 19 to (75, 100, 223.81) mm, rotated rx 2.71 ry -3.1 rz 88.36 deg; joints [-131.372, 30.115, -33.133, 91.43, 72.876, -178.92, 2497.581, -237.209, 490.363]
  MoveL 20 to (75, 200, 229.45) mm, rotated rx 2.7 ry -3.22 rz 88.36 deg; joints [-131.372, 30.326, -33.133, 91.488, 73.005, -179.133, 2397.813, -235.278, 490.363]
  MoveL 21 to (75, 300, 235.32) mm, rotated rx 8.08 ry -3.19 rz 88.2 deg; joints [-131.372, 31.343, -33.133, 96.576, 73.203, -184.409, 2304.322, -235.278, 454.993]
  MoveL 22 to (75, 400, 241.4) mm, rotated rx 8.19 ry -3.31 rz 88.18 deg; joints [-131.372, 31.625, -33.133, 96.747, 73.362, -184.784, 2204.989, -233.26, 454.993]
  MoveL 23 to (75, 500, 247.79) mm, rotated rx 9.22 ry -3.43 rz 88.13 deg; joints [-131.372, 32.415, -33.133, 97.876, 73.675, -186.401, 2108.691, -233.26, 453.753]
  MoveL 24 to (75, 600, 261.44) mm, rotated rx 23.66 ry -23.77 rz 79.03 deg; joints [-131.372, 36.733, -33.133, 102.062, 97.93, -199.637, 1868.867, -104.915, 453.752]
  MoveL 25 to (75, 700, 280.68) mm, rotated rx 20.02 ry -2.78 rz 87.99 deg; joints [-140.774, 36.733, -29.31, 107.647, 86.181, -199.637, 2042.676, -104.915, 444.348]
  MoveL 26 to (75, 800, 276.44) mm, rotated rx 22.59 ry 10.54 rz 93.42 deg; joints [-143.982, 36.733, -29.31, 113.947, 76.326, -200.447, 2102.82, -104.915, 407.634]
  MoveL 27 to (75, 900, 278.65) mm, rotated rx -15.68 ry -40.48 rz 98.44 deg; joints [-134.388, 36.733, -29.31, 82.197, 113.909, -178.747, 1521.455, 43.242, 652.984]
  Set speed (1000.0 mm/s)
  MoveL 28 to (75, 900, 278.65) mm, rotated rx -15.68 ry -40.48 rz 98.44 deg; joints [-134.388, 36.733, -29.31, 82.197, 113.909, -178.747, 1521.455, 43.242, 652.984]
  MoveL 29 to (92.55, 965.79, 205.41) mm, rotated rx -15.68 ry -40.48 rz 98.44 deg; joints [-140.37, 35.88, -29.31, 81.467, 119.907, -178.747, 1517.07, 43.241, 657.394]
  Set speed (1000.0 mm/s)
  MoveL 30 to (120.12, 805.44, 147.11) mm, rotated rx 17.49 ry -2.67 rz 88.08 deg; joints [-161.484, 35.88, -29.31, 103.644, 105.044, -192.17, 2094.235, 43.241, 495.486]
  MoveL 31 to (150, 800, 242.38) mm, rotated rx 17.49 ry -2.67 rz 88.08 deg; joints [-161.185, 35.808, -29.31, 103.678, 104.739, -192.17, 2094.235, 134.311, 524.444]
  MoveL 32 to (150, 800, 242.38) mm, rotated rx 17.49 ry -2.67 rz 88.08 deg; joints [-161.185, 35.808, -29.31, 103.678, 104.739, -192.17, 2094.235, 134.311, 524.444]
  Set speed (200.0 mm/s)
  MoveL 33 to (150, 700, 237.54) mm, rotated rx 14.66 ry -1.9 rz 88.34 deg; joints [-161.654, 33.92, -29.31, 101.832, 103.527, -189.285, 2188.918, 134.311, 524.444]
  MoveL 34 to (150, 600, 232.62) mm, rotated rx 12 ry -2.62 rz 88.21 deg; joints [-161.609, 31.991, -29.31, 99.847, 103.527, -186.551, 2266.679, 134.311, 525.169]
  MoveL 35 to (150, 500, 227.36) mm, rotated rx 11.17 ry -2.76 rz 88.2 deg; joints [-161.667, 31.223, -29.31, 99.289, 103.527, -185.506, 2359.264, 133.93, 525.169]
  MoveL 36 to (150, 400, 221.99) mm, rotated rx 13.97 ry -2.53 rz 88.19 deg; joints [-161.642, 31.223, -29.31, 101.759, 103.527, -186.378, 2461.132, 135.141, 504.462]
  MoveL 37 to (150, 300, 216.85) mm, rotated rx 13.48 ry -2.49 rz 88.21 deg; joints [-161.788, 30.69, -29.31, 101.465, 103.47, -185.658, 2557.701, 135.141, 504.462]
  MoveL 38 to (150, 200, 211.93) mm, rotated rx 12.77 ry -2.29 rz 88.27 deg; joints [-161.959, 30.018, -29.31, 101.027, 103.254, -184.725, 2654.374, 135.141, 504.462]
  MoveL 39 to (150, 100, 207.2) mm, rotated rx 12.8 ry -2.35 rz 88.25 deg; joints [-161.959, 29.816, -29.31, 101.098, 103.27, -184.532, 2752.185, 133.949, 504.462]
  MoveL 40 to (150, 0, 203.02) mm, rotated rx 12.74 ry -1.88 rz 88.36 deg; joints [-162.195, 29.772, -29.31, 101.098, 103.011, -184.412, 2857.032, 133.949, 506.753]
  Set speed (1000.0 mm/s)
  MoveL 41 to (150, 0, 203.02) mm, rotated rx 12.74 ry -1.88 rz 88.36 deg; joints [-162.195, 29.772, -29.31, 101.098, 103.011, -184.412, 2857.032, 133.949, 506.753]
  MoveL 42 to (128.05, 3.83, 105.54) mm, rotated rx 12.74 ry -1.88 rz 88.36 deg; joints [-162.291, 29.791, -29.31, 101.097, 103.109, -184.412, 2857.031, 37.709, 485.046]
  Set speed (1000.0 mm/s)
  MoveL 43 to (220.65, 4.01, 93.86) mm, rotated rx 2.55 ry -2.23 rz 88.41 deg; joints [-162.381, 29.791, -29.31, 92.09, 103.109, -181.268, 2852.075, 17.236, 664.089]
  MoveL 44 to (225, 0, 193.68) mm, rotated rx 2.55 ry -2.23 rz 88.41 deg; joints [-162.381, 29.79, -29.31, 92.09, 103.109, -181.268, 2853.288, 117.133, 668.44]
  MoveL 45 to (225, 0, 193.68) mm, rotated rx 2.55 ry -2.23 rz 88.41 deg; joints [-162.381, 29.79, -29.31, 92.09, 103.109, -181.268, 2853.288, 117.133, 668.44]
  Set speed (200.0 mm/s)
  MoveL 46 to (225, 100, 197.78) mm, rotated rx 2.48 ry -2.34 rz 88.4 deg; joints [-162.275, 29.891, -29.31, 92.001, 103.109, -181.353, 2752.783, 117.133, 667.602]
  MoveL 47 to (225, 200, 202.17) mm, rotated rx 2.48 ry -2.51 rz 88.4 deg; joints [-162.105, 29.891, -29.31, 91.999, 103.117, -181.361, 2650.435, 117.134, 664.884]
  MoveL 48 to (225, 300, 206.77) mm, rotated rx 2.74 ry -2.52 rz 88.39 deg; joints [-162.081, 30.282, -29.31, 92.128, 103.117, -181.841, 2553.676, 117.697, 664.884]
  MoveL 49 to (225, 400, 211.28) mm, rotated rx 3.42 ry -2.45 rz 88.38 deg; joints [-162.087, 30.966, -29.31, 92.575, 103.105, -182.758, 2460.23, 117.697, 664.884]
  MoveL 50 to (225, 500, 215.72) mm, rotated rx 3.72 ry -2.47 rz 88.38 deg; joints [-162.033, 31.38, -29.31, 92.737, 103.105, -183.277, 2363.307, 117.767, 664.884]
  MoveL 51 to (225, 600, 220.75) mm, rotated rx 5.54 ry -1.67 rz 88.42 deg; joints [-162.275, 32.835, -29.31, 94.068, 102.758, -185.308, 2283.425, 117.768, 664.883]
  MoveL 52 to (225, 700, 223.76) mm, rotated rx 6.11 ry -1.55 rz 88.44 deg; joints [-162.343, 33.331, -29.31, 94.465, 102.783, -185.981, 2188.915, 117.767, 663.691]
  Set speed (1000.0 mm/s)
  MoveL 53 to (225, 700, 223.76) mm, rotated rx 6.11 ry -1.55 rz 88.44 deg; joints [-162.343, 33.331, -29.31, 94.465, 102.783, -185.981, 2188.915, 117.767, 663.691]
  MoveL 54 to (214.44, 702.97, 124.36) mm, rotated rx 6.11 ry -1.55 rz 88.44 deg; joints [-162.344, 33.331, -29.31, 94.464, 102.784, -185.981, 2188.908, 18.351, 653.156]
  Set speed (1000.0 mm/s)
  MoveL 55 to (297.16, 702.27, 119.51) mm, rotated rx 1.66 ry -1.26 rz 88.45 deg; joints [-162.845, 32.919, -29.31, 90.621, 102.636, -184.182, 2188.908, 18.351, 768.606]
  MoveL 56 to (300, 700, 219.45) mm, rotated rx 1.66 ry -1.26 rz 88.45 deg; joints [-162.845, 32.919, -29.31, 90.621, 102.636, -184.182, 2188.421, 118.31, 771.407]
  MoveL 57 to (300, 700, 219.45) mm, rotated rx 1.66 ry -1.26 rz 88.45 deg; joints [-162.845, 32.919, -29.31, 90.621, 102.636, -184.182, 2188.421, 118.31, 771.407]
  Set speed (200.0 mm/s)
  MoveL 58 to (300, 600, 217.1) mm, rotated rx -0.28 ry -1.56 rz 88.44 deg; joints [-162.631, 31.395, -29.31, 89.23, 102.636, -182.032, 2271.976, 120.497, 771.408]
  MoveL 59 to (300, 500, 213.93) mm, rotated rx -0.88 ry -1.74 rz 88.44 deg; joints [-162.497, 30.775, -29.31, 88.842, 102.674, -181.213, 2364.505, 120.497, 771.408]
  MoveL 60 to (300, 400, 210.18) mm, rotated rx -0.47 ry -2.5 rz 88.45 deg; joints [-162.359, 30.775, -29.31, 89.186, 103.308, -181.34, 2457.368, 120.497, 770.637]
  MoveL 61 to (300, 300, 205.93) mm, rotated rx -1.36 ry -2.52 rz 88.46 deg; joints [-162.34, 29.951, -29.31, 88.599, 103.308, -180.217, 2549.963, 121.143, 770.638]
  MoveL 62 to (300, 200, 201.56) mm, rotated rx -1.07 ry -2.61 rz 88.46 deg; joints [-162.34, 29.932, -29.31, 88.859, 103.403, -180.287, 2649.035, 119.839, 770.638]
  MoveL 63 to (300, 100, 197.15) mm, rotated rx -0.69 ry -2.46 rz 88.45 deg; joints [-162.486, 29.932, -29.31, 89.194, 103.403, -180.408, 2751.005, 119.554, 770.123]
  MoveL 64 to (300, 0, 193.08) mm, rotated rx -2.06 ry -2.36 rz 88.47 deg; joints [-162.486, 28.762, -29.31, 88.262, 103.336, -178.782, 2841.368, 121.371, 770.126]
  Set speed (1000.0 mm/s)
  MoveL 65 to (300, 0, 193.08) mm, rotated rx -2.06 ry -2.36 rz 88.47 deg; joints [-162.486, 28.762, -29.31, 88.262, 103.336, -178.782, 2841.368, 121.371, 770.126]
  MoveL 66 to (303.7, 4.02, 93.23) mm, rotated rx -2.06 ry -2.36 rz 88.47 deg; joints [-162.486, 28.762, -29.31, 88.262, 103.336, -178.782, 2839.932, 21.451, 773.819]
  Set speed (1000.0 mm/s)
  MoveL 67 to (382.7, 3.94, 97.57) mm, rotated rx -4.36 ry -2.38 rz 88.5 deg; joints [-162.412, 28.762, -29.31, 86.236, 103.336, -178.068, 2837.249, 25.97, 872.373]
  MoveL 68 to (375, 0, 197.2) mm, rotated rx -4.36 ry -2.38 rz 88.5 deg; joints [-162.412, 28.762, -29.31, 86.236, 103.336, -178.068, 2838.719, 125.661, 864.677]
  MoveL 69 to (375, 0, 197.2) mm, rotated rx -4.36 ry -2.38 rz 88.5 deg; joints [-162.412, 28.762, -29.31, 86.236, 103.336, -178.068, 2838.719, 125.661, 864.677]
  Set speed (200.0 mm/s)
  MoveL 70 to (375, 100, 201.22) mm, rotated rx -4.3 ry -2.5 rz 88.51 deg; joints [-162.336, 29.015, -29.31, 86.228, 103.366, -178.339, 2739.592, 125.662, 864.558]
  MoveL 71 to (375, 200, 205.44) mm, rotated rx -4.44 ry -2.52 rz 88.51 deg; joints [-162.318, 29.145, -29.31, 86.081, 103.366, -178.429, 2640.442, 126.742, 864.557]
  MoveL 72 to (375, 300, 209.49) mm, rotated rx -3.68 ry -2.33 rz 88.49 deg; joints [-162.457, 29.879, -29.31, 86.564, 103.249, -179.426, 2549.304, 126.742, 864.556]
  MoveL 73 to (375, 400, 213.08) mm, rotated rx -3.23 ry -2.01 rz 88.46 deg; joints [-162.601, 30.402, -29.31, 86.837, 103.043, -180.109, 2457.26, 126.742, 864.556]
  MoveL 74 to (375, 500, 216.05) mm, rotated rx -2.67 ry -1.73 rz 88.45 deg; joints [-162.789, 30.998, -29.31, 87.195, 102.922, -180.903, 2365.744, 126.742, 864.556]
  MoveL 75 to (375, 600, 218.52) mm, rotated rx -1.86 ry -1.36 rz 88.43 deg; joints [-163.06, 31.755, -29.31, 87.734, 102.806, -181.932, 2276.656, 126.742, 864.555]
  Set speed (1000.0 mm/s)
  MoveL 76 to (375, 600, 218.52) mm, rotated rx -1.86 ry -1.36 rz 88.43 deg; joints [-163.06, 31.755, -29.31, 87.734, 102.806, -181.932, 2276.656, 126.742, 864.555]
  MoveL 77 to (378.31, 602.28, 118.6) mm, rotated rx -1.86 ry -1.36 rz 88.43 deg; joints [-163.06, 31.719, -29.31, 87.742, 102.807, -181.895, 2276.656, 26.893, 867.444]
  Set speed (1000.0 mm/s)
  MoveL 78 to (454.83, 601.84, 122) mm, rotated rx -2.74 ry -1.13 rz 88.42 deg; joints [-163.06, 31.69, -29.31, 86.972, 102.556, -181.6, 2276.657, 29.818, 951.2]
  MoveL 79 to (450, 600, 221.87) mm, rotated rx -2.74 ry -1.13 rz 88.42 deg; joints [-163.06, 31.773, -29.31, 86.954, 102.551, -181.685, 2276.656, 129.48, 947.372]
  MoveL 80 to (450, 600, 221.87) mm, rotated rx -2.74 ry -1.13 rz 88.42 deg; joints [-163.06, 31.773, -29.31, 86.954, 102.551, -181.685, 2276.656, 129.48, 947.372]
  Set speed (200.0 mm/s)
  MoveL 81 to (450, 500, 220.16) mm, rotated rx -3.81 ry -0.92 rz 88.4 deg; joints [-163.06, 30.826, -29.31, 86.215, 102.377, -180.396, 2370.308, 132.655, 947.373]
  MoveL 82 to (450, 400, 218.21) mm, rotated rx -4.34 ry -1.74 rz 88.45 deg; joints [-162.66, 30.264, -29.31, 85.883, 102.838, -179.631, 2456.489, 132.655, 947.374]
  MoveL 83 to (450, 300, 215.34) mm, rotated rx -4.61 ry -1.94 rz 88.47 deg; joints [-162.526, 29.864, -29.31, 85.74, 102.939, -179.129, 2550.615, 132.655, 947.374]
  MoveL 84 to (450, 200, 211.78) mm, rotated rx -4.24 ry -2.17 rz 88.48 deg; joints [-162.526, 29.864, -29.31, 86.077, 103.169, -179.244, 2648.628, 132.472, 946.812]
  MoveL 85 to (450, 100, 207.82) mm, rotated rx -4.65 ry -2.42 rz 88.51 deg; joints [-162.426, 29.366, -29.31, 85.837, 103.362, -178.599, 2741.604, 132.472, 946.812]
  MoveL 86 to (450, 0, 203.99) mm, rotated rx -4.99 ry -2.31 rz 88.5 deg; joints [-162.431, 28.907, -29.31, 85.643, 103.291, -178.024, 2838.512, 132.472, 946.812]
  Set speed (1000.0 mm/s)
  MoveL 87 to (450, 0, 203.99) mm, rotated rx -4.99 ry -2.31 rz 88.5 deg; joints [-162.431, 28.907, -29.31, 85.643, 103.291, -178.024, 2838.512, 132.472, 946.812]
  MoveL 88 to (458.8, 3.78, 104.45) mm, rotated rx -4.99 ry -2.31 rz 88.5 deg; joints [-162.431, 28.907, -29.31, 85.643, 103.291, -178.024, 2837.167, 32.868, 955.604]
  Set speed (1000.0 mm/s)
  MoveL 89 to (515.12, 3.49, 104.06) mm, rotated rx 5.73 ry -1.85 rz 88.41 deg; joints [-162.551, 28.907, -29.31, 95.108, 102.904, -181.329, 2840.382, 32.868, 920.358]
  MoveL 90 to (525, 0, 203.5) mm, rotated rx 5.73 ry -1.85 rz 88.41 deg; joints [-162.551, 28.907, -29.31, 95.108, 102.904, -181.329, 2840.929, 132.377, 930.229]
  MoveL 91 to (525, 0, 203.5) mm, rotated rx 5.73 ry -1.85 rz 88.41 deg; joints [-162.551, 28.907, -29.31, 95.108, 102.904, -181.329, 2840.929, 132.377, 930.229]
  Set speed (200.0 mm/s)
  MoveL 92 to (525, 100, 207.22) mm, rotated rx 5.48 ry -2.06 rz 88.39 deg; joints [-162.441, 28.953, -29.31, 94.874, 103.008, -181.312, 2738.998, 132.377, 930.229]
  MoveL 93 to (525, 200, 211.32) mm, rotated rx 5.33 ry -2.41 rz 88.36 deg; joints [-162.259, 28.983, -29.31, 94.718, 103.169, -181.312, 2635.468, 132.377, 929.32]
  MoveL 94 to (525, 300, 215.9) mm, rotated rx 5.32 ry -2.56 rz 88.34 deg; joints [-162.095, 29.055, -29.31, 94.686, 103.169, -181.397, 2533.967, 132.377, 927.595]
  MoveL 95 to (525, 400, 220.62) mm, rotated rx 3.08 ry -2.6 rz 88.38 deg; joints [-162.094, 29.055, -29.31, 92.712, 103.169, -180.69, 2433.601, 133.162, 943.953]
  MoveL 96 to (525, 500, 224.64) mm, rotated rx 0.01 ry -1.71 rz 88.44 deg; joints [-162.302, 29.055, -29.31, 90.017, 102.478, -179.724, 2342.137, 133.162, 967.298]
  Set speed (1000.0 mm/s)
  MoveL 97 to (525, 500, 224.64) mm, rotated rx 0.01 ry -1.71 rz 88.44 deg; joints [-162.302, 29.055, -29.31, 90.017, 102.478, -179.724, 2342.137, 133.162, 967.298]
  MoveL 98 to (525.06, 502.99, 124.68) mm, rotated rx 0.01 ry -1.71 rz 88.44 deg; joints [-162.302, 29.055, -29.31, 90.017, 102.478, -179.724, 2341.831, 33.165, 967.376]

